(* IEC 61131-3 sources: daoli-st-library/DL_Process (part 7) *)

(* ---- FB_DL_SplicerAutoJoint.st ---- *)
//==============================================================================
// 功能块：FB_DL_SplicerAutoJoint ｜ 中文名称：自动接膜零停机顺控
// 所属子库：DL_Process ｜ 版本：v1.1.1 ｜ 兼容：CODESYS V3.5+ / TwinCAT 3 / 汇川 InoProShop
// 功能描述：卷材设备自动接膜（零停机换卷）顺控：旧卷余量预警 → 新卷预加速 → 速度同步
//           确认（容差 + 保持时长双条件）→ 裁切压合 → 尾料处理 → 回到监测相。
//           安全铁律：未同步绝不裁切——速度差超容差或保持时长不足时裁切一律挂起，宁可
//           等，不裁切（拉断料带的代价远高于停一拍）。余量按面积（卷径平方）比例折算，
//           按直径线性折算会把余量算大一倍以上（量纲教训：卷材体积随直径平方变化）。
//           本件只发预加速/裁切指令与状态，不驱动伺服、不控气阀（执行器归设备层）。
// 开源溯源 (Origin)：道莅 clean-room 防御性实现（原创，参考 公开工程惯例 分类与参数域）
// 单位表：卷径/芯径/满卷直径[mm] / 线速度[米每分] / 余量与预警门限[百分数] /
//         同步容差[百分数] / 时间窗[ms] / 扫描间隔[ms] / 接膜次数[次]
// 错误码表：16#0005_040A 信息级（余量预警触发，上升沿一次，不置 bError）/
//           16#0005_040B 信息级（同步窗未达，裁切挂起，不置 bError）/ 16#0005_0351
//           故障级（预加速超时中止且不裁切；兼「卷径组态非法（满卷直径 ≤ 芯径）」组态
//           分支，映射见本行反证句）/ 16#0005_0352 故障级（胶带未就绪或刀未归零，禁止
//           接膜，置 bError + 撤全部指令）/ 16#0005_0353 故障级（输入非有限，以及状态机
//           ELSE 非法状态兜底）。0351 共用反证句：组态非法、预加速超时与同步相超时
//           （v1.1.0 新增）在现有输出组合下不可观测出差异（均为 bError + bPreAccelCmd 撤
//           + bCutCmd 撤 + bSyncOk 撤 + bValid 撤），同步超时另由 bSyncTimeout 单拍事件可区分观测；
//           §4.17 亦明示组态分支映射入 0351，故共用不越段。0353 共用反证句：非有限
//           输入与非法状态在输出上同为全撤 + bError + eFault，不可观测出差异，故共用。
// 状态机：E_DL_SplicerState（eIdle=0 待机 / eMonitor=10 余量监测 / ePreAccel=20 新卷
//           预加速 / eSyncWait=30 同步确认 / eJointing=40 裁切压合 / eFault=99 故障兜底），
//           CASE 含 ELSE 兜底，ELSE 置 0353 且撤全部指令、许可撤。
// 边界行为：① 余量按面积比例 ((D^2 − core^2)/(full^2 − core^2)) x 100，D 低于芯径钳 0、
//           高于满卷钳 100；② fFullDiaMm <= fCoreDiaMm → 故障 0351 组态分支（分母为零
//           会产出伪余量，先判后算）；③ 预加速超 tPreAccelMax → 故障 0351 + 中止且绝不
//           裁切（停机保料优于拉断）；④ 同步未达（速度差 > 容差，或保持不足 tSyncHold）
//           → 裁切挂起 + 信息 040B（安全侧：宁可等，不裁切）；⑤ bTapeOk 或 bKnifeHome
//           为 FALSE → 禁止接膜 + 故障 0352；⑥ bStop → 中止并回 eIdle（同③不裁切）；
//           ⑦ 余量预警上升沿 → 信息 040A（用沿检测，防每拍刷屏）。
// 修订历史：v1.0.0 2026-11-17 首版（R25 派单 · §4.17）
//           v1.0.1 2026-11-17 终审补 eSyncWait 的「进相前置消失」第二退出条件（对外引脚契约零变更）：
//           bNewRollReady 撤销时退回 ePreAccel 相，由 tPreAccelMax 超时闸兜住，避免 bPreAccelCmd
//           长期拉住空卷（R98 家族）。两相 bCutCmd 均为 FALSE，「未同步绝不裁切」铁律不受影响。
//           v1.1.0 2026-11-17 R27 欠账收口（MINOR 升级，引脚契约只增不改、既有码位零变更）：
//           eSyncWait 相新增引脚 tSyncMax（同步等待超时，默认 T#5S）与自有计时器 fbTonSyncMax
//           （每周期无条件调用，仅 IN 条件化）；速度差持续超容差达 tSyncMax 即复用故障级 0351
//           （同段共用，反证句见错误码表 0351 行）并中止，bCutCmd 全程保持 FALSE；新增输出
//           bSyncTimeout（超时单拍事件，供审计计数）。
//           原挂账 R112 三要素收口：复现条件 = bNewRollReady 保持 TRUE 而速度差持续超容差（旧版将
//           无限期停在同步相）；禁用范围 = 无人值守连续线未配该超时者不得无人看管运行；修法取
//           ①新增 tSyncMax 引脚（默认 5 s 从紧口径）。
//           验收向量（VERSION 修订记录同步登记）：新卷就绪后速度差恒定 5%、容差 2% →
//           tSyncMax 之后置 0351、bSyncTimeout 单拍 TRUE、bCutCmd 全程 FALSE。
//           v1.1.1 2026-11-17 R27 终审修复（对外引脚与码位零变更）：fbTonSyncMax 的 IN 由
//           「eSyncWait AND NOT bSpeedWithin」改为「eSyncWait」按相驻留计时。原实现的看门狗
//           只在速度差超出容差时累积：速度差在容差边界抖动（模拟量噪声常态）时，同步超时
//           计时器与同步保持计时器交替复位，两者永不完成 → 相内无限滞留、段 8B 永不触发，
//           bPreAccelCmd 长期拉住空卷，恰是 v1.1.0 要收口的故障模式在抖动输入下的复现。
//           改为按相驻留计时后，相内总等待时长有上界，抖动亦能收口；正常同步（远早于
//           tSyncMax 完成）行为不变。验收向量：速度差在 2% 容差上下逐拍抖动 → tSyncMax 后 0351。
//==============================================================================
(*------------------------------------------------------------------------------
 * 枚举: E_DL_SplicerState（归属 DL_Process，与 FB_DL_SplicerAutoJoint 同文件）
 *----------------------------------------------------------------------------*)
TYPE E_DL_SplicerState :
(
    eIdle     := 0,   // 待机：指令全撤 / Idle, every command dropped
    eMonitor  := 10,  // 余量监测：算余量、报预警 / Monitoring the remaining roll
    ePreAccel := 20,  // 预加速：新卷升速，等就绪与同步 / Pre-accelerating the new roll
    eSyncWait := 30,  // 同步确认：速度差在容差内且保持达时 / Confirming the speed match
    eJointing := 40,  // 裁切压合：出裁切指令并在接膜窗内完成 / Cutting and joining
    eFault    := 99   // 故障兜底：超时/胶带刀具不就绪/非有限/非法状态 / Fault fallback
);
END_TYPE

(*==============================================================================
 * 功能块: FB_DL_SplicerAutoJoint
 * 调用约定: 每个扫描周期无条件调用一次；uDeltaTimeMs 必须注入真实任务间隔。
 *============================================================================*)
FUNCTION_BLOCK FB_DL_SplicerAutoJoint
VAR_INPUT
    fUnwindDiaMm    : LREAL;                       // 旧卷当前卷径 [mm] / Current unwinding roll diameter [mm]
    fCoreDiaMm      : LREAL;                       // 芯径 [mm]，须 > 0 / Core diameter [mm], must be > 0
    fFullDiaMm      : LREAL;                       // 满卷直径 [mm]，须 > 芯径 / Full roll diameter [mm], must exceed the core
    fWebSpeedMpm    : LREAL;                       // 旧卷线速度 [米每分] / Current web speed [m per min]
    fNewRollSpeedMpm : LREAL;                      // 新卷表面线速度 [米每分] / New roll surface speed [m per min]
    fRemainWarnPct  : LREAL := 15.0;               // 余量预警门限 [百分数] / Remaining-roll warning threshold [percent]
    fSyncTolPct     : LREAL := 2.0;                // 速度同步容差 [百分数] / Speed match tolerance [percent]
    tSyncHold       : TIME := T#500MS;             // 同步保持确认时长 [ms] / Speed match hold time [ms]
    tPreAccelMax    : TIME := T#20S;               // 预加速超时 [ms] / Pre-acceleration timeout [ms]
    tJointMax       : TIME := T#5S;                // 接膜（裁切压合）窗 [ms] / Joint window [ms]
    tSyncMax        : TIME := T#5S;                // 同步等待超时 [ms]，默认 5 s（eSyncWait 自有看门狗，小于 1 s 钳 1 s）/ Sync wait timeout [ms]
    bNewRollReady   : BOOL;                        // 新卷就绪（装卷到位、气路正常）/ New roll ready
    bKnifeHome      : BOOL;                        // 切刀在零位 / Knife at home position
    bTapeOk         : BOOL;                        // 胶带就绪 / Tape ready
    bStart          : BOOL;                        // 启动（取上升沿）/ Start, rising edge
    bStop           : BOOL;                        // 停止（中止并回待机，绝不裁切）/ Stop, aborts without cutting
    bReset          : BOOL;                        // 复位，上升沿回待机并清故障 / Reset, rising edge returns to idle
    uDeltaTimeMs    : UDINT;                       // 扫描间隔 [ms]，调用方注入，禁系统时间函数 / Scan interval [ms], caller-injected
END_VAR
VAR_OUTPUT
    bWarnLowRoll    : BOOL;                        // 余量预警（电平）/ Low-roll warning, level
    bPreAccelCmd    : BOOL;                        // 新卷预加速指令 / Pre-acceleration command
    bSyncOk         : BOOL;                        // 速度同步确认（容差 + 保持时长双条件）/ Speed match confirmed
    bSyncTimeout    : BOOL;                        // 同步超时事件（单拍脉冲，v1.1.0 新增）/ Sync-timeout event, single-scan pulse
    bCutCmd         : BOOL;                        // 裁切指令（未同步绝不为 TRUE）/ Cut command, never TRUE unless matched
    bJointDone      : BOOL;                        // 接膜完成（单拍脉冲）/ Joint completed, single-scan pulse
    fRemainPct      : LREAL;                       // 旧卷余量 [百分数]，按面积比例 / Remaining roll [percent], by area ratio
    uJointCount     : UDINT;                       // 接膜次数 [次]，饱和 / Joint count [pcs], saturating
    eErr            : UDINT;                       // 错误码，0 = 无错，码位 16#0005_040A 起信息级、16#0005_0351 起故障级（分带见错误码表） / Error code, 0 = no error, band info/fault per the code table
    bError          : BOOL;                        // 故障级标志，仅故障级错误置位 / Fault-class flag, set only on fault-level codes
    bValid          : BOOL;                        // 状态输出可用标志，失能/故障闸显式 FALSE / Status usable flag, explicit FALSE on disable/fault gates
    eState          : E_DL_SplicerState;           // 主状态机当前状态 / Current state of the main state machine
END_VAR
VAR
    fbReset         : R_TRIG;                      // 复位上升沿检测实例 / Reset rising edge detector
    fbStart         : R_TRIG;                      // 启动上升沿检测实例 / Start rising edge detector
    fbWarn          : R_TRIG;                      // 余量预警上升沿检测实例 / Low-roll warning rising edge detector
    fbTonPreAccel   : TON;                         // 预加速超时定时器实例 / Pre-acceleration timeout timer
    fbTonSyncHold   : TON;                         // 同步保持定时器实例 / Speed match hold timer
    fbTonJoint      : TON;                         // 接膜窗定时器实例 / Joint window timer
    fbTonSyncMax    : TON;                         // 同步相自有超时定时器实例（每周期无条件调用）/ Sync-phase watchdog timer instance
    tSyncMaxUse     : TIME;                        // 生效同步超时（下限钳 1 s 防误配置）/ Effective sync timeout, floored at 1 s
    fCoreSqMm2      : LREAL;                       // 芯径平方 [平方毫米] / Core diameter squared [mm2]
    fFullSqMm2      : LREAL;                       // 满卷直径平方 [平方毫米] / Full diameter squared [mm2]
    fDenomMm2       : LREAL;                       // 面积分母（满卷平方 − 芯径平方）[平方毫米] / Area denominator [mm2]
    fRemainNumMm2   : LREAL;                       // 面积分子（当前平方 − 芯径平方）[平方毫米] / Area numerator [mm2]
    fSpeedDiffPct   : LREAL;                       // 新旧卷速度差 [百分数] / Speed difference [percent]
    fTolEffPct      : LREAL;                       // 生效同步容差 [百分数] / Effective sync tolerance [percent]
    fWarnEffPct     : LREAL;                       // 生效预警门限 [百分数] / Effective warning threshold [percent]
    bNonFin         : BOOL;                        // 非有限判定中间标志 / Non-finite detection intermediate flag
    bSpeedWithin    : BOOL;                        // 速度差在容差内（瞬时）/ Speed difference within tolerance, instantaneous
    bJointOk        : BOOL;                        // 胶带与刀具均就绪 / Tape and knife both ready
    bFirstScan      : BOOL := TRUE;                // 上电首拍标志 / First-scan flag
END_VAR
VAR CONSTANT
    DL_SPJ_CODE_INFO_1 : UDINT := 16#0005_040A;    // 信息级槽 1（余量预警触发） / info slot 1
    DL_SPJ_CODE_INFO_2 : UDINT := 16#0005_040B;    // 信息级槽 2（同步窗未达，裁切挂起） / info slot 2
    DL_SPJ_CODE_FLT_1  : UDINT := 16#0005_0351;    // 故障级槽 1（预加速超时/卷径组态非法） / fault slot 1
    DL_SPJ_CODE_FLT_2  : UDINT := 16#0005_0352;    // 故障级槽 2（胶带未就绪/刀未归零） / fault slot 2
    DL_SPJ_CODE_FLT_3  : UDINT := 16#0005_0353;    // 故障级槽 3（非有限/非法状态兜底） / fault slot 3
    DL_SPJ_CNT_MAX     : UDINT := 16#FFFF_FFFE;    // 接膜计数饱和值 [次] / Joint counter saturation
    DL_SPJ_PCT         : LREAL := 100.0;           // 百分数系数 [百分数] / Percent factor
    DL_SPJ_ZERO        : LREAL := 0.0;             // 零值常量，避免裸字面量 [—] / Zero constant, avoids a bare literal
    DL_SPJ_TOL         : LREAL := 1.0E-6;          // 浮点比较容差 [—] / Float comparison tolerance
    DL_SPJ_INF         : LREAL := 1.7976931348623157E308; // LREAL 幅值上限，Inf 判据 / LREAL magnitude ceiling
END_VAR

(*------------------------------------------------------------------------------
 * 段 1｜无条件刷新区（红线 5）：三条沿检测与三个定时器在任意分支之外周期调用；
 *       定时器 IN 取上拍状态（单拍滞后对秒级时间窗无影响），计时链永不断流
 *----------------------------------------------------------------------------*)
bJointDone := FALSE;                               // 接膜完成为单拍脉冲，逐拍先清 / single-scan pulse cleared first
bSyncTimeout := FALSE;                             // 同步超时为单拍事件，逐拍先清 / sync-timeout event cleared first
tSyncMaxUse := tSyncMax;                           // 生效超时取引脚值 / effective timeout from the pin
IF tSyncMaxUse < T#1S THEN
    tSyncMaxUse := T#1S;                           // 超时下限钳 1 s（防 0 配置入相同拍误报）/ floored at 1 s
END_IF
fbReset(CLK := bReset);                            // 复位沿检测无条件刷新 / reset edge refreshed unconditionally
fbStart(CLK := bStart);                            // 启动沿检测无条件刷新 / start edge refreshed unconditionally
fbTonPreAccel(IN := (eState = E_DL_SplicerState.ePreAccel), PT := tPreAccelMax);   // 预加速超时计时 / pre-acceleration timeout
fbTonSyncHold(IN := (eState = E_DL_SplicerState.eSyncWait) AND bSpeedWithin, PT := tSyncHold);   // 同步保持计时 / speed match hold
fbTonJoint(IN := (eState = E_DL_SplicerState.eJointing), PT := tJointMax);         // 接膜窗计时 / joint window
fbTonSyncMax(IN := (eState = E_DL_SplicerState.eSyncWait), PT := tSyncMaxUse);   // v1.1.1 改为按相驻留计时（见修订史 R27-3）/ sync watchdog on phase residency
fbWarn(CLK := bWarnLowRoll);                       // 预警上升沿检测无条件刷新 / warning edge refreshed unconditionally

(*------------------------------------------------------------------------------
 * 段 2｜复位沿处理（改写置于沿后，防吞沿 R39）
 *----------------------------------------------------------------------------*)
IF fbReset.Q THEN
    eState := E_DL_SplicerState.eIdle;
    eErr   := 0;                        // 复位清码 / reset clears the code
    bError := FALSE;                               // 复位清故障 / reset clears the fault
    bPreAccelCmd := FALSE;                         // 预加速指令撤 / pre-acceleration dropped
    bCutCmd := FALSE;                              // 裁切指令撤 / cut command dropped
    bSyncOk := FALSE;                              // 同步确认撤 / sync confirmation dropped
    bFirstScan := TRUE;                            // 重新首拍化 / re-initialize first scan
END_IF

(*------------------------------------------------------------------------------
 * 段 3｜非有限输入闸：映射入 0353（与非法状态共用，反证句见错误码表）
 *       安全侧：撤全部指令，绝不裁切
 *----------------------------------------------------------------------------*)
bNonFin := (fUnwindDiaMm <> fUnwindDiaMm) OR (ABS(fUnwindDiaMm) >= DL_SPJ_INF)
        OR (fCoreDiaMm <> fCoreDiaMm) OR (ABS(fCoreDiaMm) >= DL_SPJ_INF)
        OR (fFullDiaMm <> fFullDiaMm) OR (ABS(fFullDiaMm) >= DL_SPJ_INF)
        OR (fWebSpeedMpm <> fWebSpeedMpm) OR (ABS(fWebSpeedMpm) >= DL_SPJ_INF)
        OR (fNewRollSpeedMpm <> fNewRollSpeedMpm) OR (ABS(fNewRollSpeedMpm) >= DL_SPJ_INF)
        OR (fRemainWarnPct <> fRemainWarnPct) OR (ABS(fRemainWarnPct) >= DL_SPJ_INF)
        OR (fSyncTolPct <> fSyncTolPct) OR (ABS(fSyncTolPct) >= DL_SPJ_INF);   // 引脚非有限汇总 / pins non-finite
IF bNonFin THEN
    eState := E_DL_SplicerState.eFault;            // 进故障相 / enter fault state
    eErr   := DL_SPJ_CODE_FLT_3;                   // 故障级：输入非有限 / fault: non-finite input
    bError := TRUE;                                // 故障级必置 bError（R45 配对）/ fault-class pairs with bError
    bValid := FALSE;                               // 状态不可用 / status unusable
    bPreAccelCmd := FALSE;                         // 预加速指令撤 / pre-acceleration dropped
    bCutCmd := FALSE;                              // 裁切指令撤（安全侧：绝不裁切）/ cut dropped, never cut
    bSyncOk := FALSE;                              // 同步确认撤 / sync confirmation dropped
    RETURN;
END_IF

(*------------------------------------------------------------------------------
 * 段 4｜卷径组态闸：满卷直径必须严格大于芯径（否则面积分母为零，余量必假）
 *       §4.17 明示本组态分支映射入 0351
 *----------------------------------------------------------------------------*)
IF (fCoreDiaMm <= DL_SPJ_TOL) OR (fFullDiaMm <= fCoreDiaMm + DL_SPJ_TOL) THEN
    eState := E_DL_SplicerState.eFault;            // 进故障相 / enter fault state
    eErr   := DL_SPJ_CODE_FLT_1;                   // 故障级：卷径组态非法（映射入 0351）/ fault: roll diameter configuration invalid
    bError := TRUE;                                // 故障级必置 bError（R45 配对）/ fault-class pairs with bError
    bValid := FALSE;                               // 状态不可用 / status unusable
    bPreAccelCmd := FALSE;                         // 预加速指令撤 / pre-acceleration dropped
    bCutCmd := FALSE;                              // 裁切指令撤安全侧 / cut dropped, safe side
    bSyncOk := FALSE;                              // 同步确认撤 / sync confirmation dropped
    fRemainPct := DL_SPJ_ZERO;                     // 余量不可算，输出 0 而不是伪值 / remaining reported as 0, not a fake value
    RETURN;
END_IF

(*------------------------------------------------------------------------------
 * 段 5｜余量面积比例折算：((D^2 − core^2) / (full^2 − core^2)) x 100
 *       按直径线性折算会把余量算大一倍以上（面积随直径平方变化，R12 同族量纲教训）
 *----------------------------------------------------------------------------*)
fCoreSqMm2 := fCoreDiaMm * fCoreDiaMm;             // 芯径平方 [平方毫米] / core squared [mm2]
fFullSqMm2 := fFullDiaMm * fFullDiaMm;             // 满卷直径平方 [平方毫米] / full squared [mm2]
fDenomMm2 := fFullSqMm2 - fCoreSqMm2;              // 面积分母（段 4 已保证为正）[平方毫米] / area denominator, proven positive
fRemainNumMm2 := (fUnwindDiaMm * fUnwindDiaMm) - fCoreSqMm2;   // 面积分子 [平方毫米] / area numerator [mm2]
IF fRemainNumMm2 < DL_SPJ_ZERO THEN
    fRemainNumMm2 := DL_SPJ_ZERO;                  // 卷径低于芯径：分子钳零（欠卷异常不产出负余量）/ numerator floored at zero
END_IF
fRemainPct := fRemainNumMm2 / fDenomMm2 * DL_SPJ_PCT;   // 余量 [百分数] / remaining [percent]
IF fRemainPct > DL_SPJ_PCT THEN
    fRemainPct := DL_SPJ_PCT;                      // 卷径超满卷：钳 100 / clamped to 100
END_IF
IF fRemainPct < DL_SPJ_ZERO THEN
    fRemainPct := DL_SPJ_ZERO;                     // 下限防护 / floor guard
END_IF
fWarnEffPct := fRemainWarnPct;                     // 预警门限工作副本 [百分数] / warning threshold working copy
IF fWarnEffPct < DL_SPJ_ZERO THEN
    fWarnEffPct := DL_SPJ_ZERO;                    // 门限下限钳位 / threshold floored
END_IF
IF fWarnEffPct > DL_SPJ_PCT THEN
    fWarnEffPct := DL_SPJ_PCT;                     // 门限上限钳位 / threshold clamped to 100
END_IF
bWarnLowRoll := (fRemainPct <= fWarnEffPct);       // 余量预警（电平）/ low-roll warning, level

(*------------------------------------------------------------------------------
 * 段 6｜速度同步判据：|旧卷 − 新卷| / 旧卷 x 100 <= 容差（除子先判零，低速记不同步）
 *----------------------------------------------------------------------------*)
fTolEffPct := fSyncTolPct;                         // 容差工作副本 [百分数] / tolerance working copy
IF fTolEffPct < DL_SPJ_ZERO THEN
    fTolEffPct := DL_SPJ_ZERO;                     // 负容差钳零（等价于要求完全相等）/ negative tolerance floored
END_IF
IF fWebSpeedMpm > DL_SPJ_TOL THEN
    fSpeedDiffPct := ABS(fWebSpeedMpm - fNewRollSpeedMpm) / fWebSpeedMpm * DL_SPJ_PCT;   // 速度差 [百分数] / speed difference [percent]
    bSpeedWithin := (fSpeedDiffPct <= fTolEffPct); // 容差内判据 / within-tolerance predicate
ELSE
    fSpeedDiffPct := DL_SPJ_PCT;                   // 旧卷静止：速度差按满刻度记（不可判即不同步）/ web at standstill, treated as not matched
    bSpeedWithin := FALSE;                         // 静止时不允许裁切 / no cut while the web stands still
END_IF
bJointOk := bTapeOk AND bKnifeHome;                // 胶带与刀具就绪判据 / tape and knife ready predicate
bSyncOk := bSpeedWithin AND fbTonSyncHold.Q AND (eState = E_DL_SplicerState.eSyncWait);   // 同步确认＝容差内且保持达时 / match confirmed

(*------------------------------------------------------------------------------
 * 段 7｜禁止接膜闸：胶带未就绪或刀未归零 → 0352 + 撤指令（不裁切）
 *----------------------------------------------------------------------------*)
IF (NOT bJointOk) AND ((eState = E_DL_SplicerState.ePreAccel) OR (eState = E_DL_SplicerState.eSyncWait)
                       OR (eState = E_DL_SplicerState.eJointing)) THEN
    eState := E_DL_SplicerState.eFault;            // 进故障相 / enter fault state
    eErr   := DL_SPJ_CODE_FLT_2;                   // 故障级：胶带未就绪/刀未归零，禁止接膜 / fault: tape or knife not ready
    bError := TRUE;                                // 故障级必置 bError（R45 配对）/ fault-class pairs with bError
    bValid := FALSE;                               // 状态不可用 / status unusable
    bPreAccelCmd := FALSE;                         // 预加速指令撤 / pre-acceleration dropped
    bCutCmd := FALSE;                              // 裁切指令撤（禁止接膜）/ cut dropped, joining forbidden
    bSyncOk := FALSE;                              // 同步确认撤 / sync confirmation dropped
    RETURN;
END_IF

(*------------------------------------------------------------------------------
 * 段 8｜预加速超时闸：0351 + 中止且绝不裁切（停机保料优于拉断）
 *----------------------------------------------------------------------------*)
IF (eState = E_DL_SplicerState.ePreAccel) AND fbTonPreAccel.Q THEN
    eState := E_DL_SplicerState.eFault;            // 进故障相 / enter fault state
    eErr   := DL_SPJ_CODE_FLT_1;                   // 故障级：预加速超时，中止且不裁切 / fault: pre-acceleration timeout, abort without cutting
    bError := TRUE;                                // 故障级必置 bError（R45 配对）/ fault-class pairs with bError
    bValid := FALSE;                               // 状态不可用 / status unusable
    bPreAccelCmd := FALSE;                         // 预加速指令撤 / pre-acceleration dropped
    bCutCmd := FALSE;                              // 裁切指令撤（绝不裁切）/ cut dropped, never cut
    bSyncOk := FALSE;                              // 同步确认撤 / sync confirmation dropped
    RETURN;
END_IF

(*------------------------------------------------------------------------------
 * 段 8B｜同步相超时闸（v1.1.0 欠账收口，R112 家族）：速度差持续超容差达 tSyncMax
 *       → 复用故障级 0351 并中止，bCutCmd 全程 FALSE（安全铁律：未同步绝不裁切）
 *----------------------------------------------------------------------------*)
IF (eState = E_DL_SplicerState.eSyncWait) AND fbTonSyncMax.Q THEN
    eState := E_DL_SplicerState.eFault;            // 进故障相 / enter fault state
    eErr   := DL_SPJ_CODE_FLT_1;                   // 故障级：同步超时（与预加速超时同段共用，反证句见头注）/ fault: sync timeout
    bError := TRUE;                                // 故障级必置 bError（R45 配对）/ fault-class pairs with bError
    bValid := FALSE;                               // 状态不可用 / status unusable
    bPreAccelCmd := FALSE;                         // 预加速指令撤 / pre-acceleration dropped
    bCutCmd := FALSE;                              // 裁切指令撤（绝不裁切）/ cut dropped, never cut
    bSyncOk := FALSE;                              // 同步确认撤 / sync confirmation dropped
    bSyncTimeout := TRUE;                          // 同步超时单拍事件 / single-scan sync-timeout event
    RETURN;
END_IF

(*------------------------------------------------------------------------------
 * 段 9｜状态机：CASE 含 ELSE 兜底（非法状态 → 0353 + 撤全部指令 + 许可撤）
 *----------------------------------------------------------------------------*)
CASE eState OF

    E_DL_SplicerState.eIdle:
        bPreAccelCmd := FALSE;                     // 待机预加速撤 / pre-acceleration dropped in idle
        bCutCmd := FALSE;                          // 待机裁切撤 / cut dropped in idle
        bSyncOk := FALSE;                          // 待机同步确认撤 / sync confirmation dropped in idle
        bValid := FALSE;                           // 失能闸显式不可用（R72）/ explicit FALSE on the disable gate
        eErr := 0;                      // 待机无错 / no error in idle
        bError := FALSE;                           // 待机无故障 / no fault in idle
        IF fbStart.Q THEN
            IF bJointOk THEN
                eState := E_DL_SplicerState.ePreAccel;   // 就绪才允许预加速 / pre-acceleration only when ready
                bFirstScan := FALSE;               // 首拍标志清除 / first-scan flag cleared
            ELSE
                eState := E_DL_SplicerState.eFault;      // 不就绪直接进故障相（0352）/ not ready enters the fault state
                eErr := DL_SPJ_CODE_FLT_2;         // 故障级：胶带未就绪/刀未归零 / fault: tape or knife not ready
                bError := TRUE;                    // 故障级必置 bError（R45 配对）/ fault-class pairs with bError
            END_IF
        ELSE
            eState := E_DL_SplicerState.eMonitor;  // 无启动沿：进常驻余量监测相（监测是被动功能，无需启动）/ passive monitoring needs no start
        END_IF

    E_DL_SplicerState.eMonitor:
        bPreAccelCmd := FALSE;                     // 监测相不预加速 / no pre-acceleration while monitoring
        bCutCmd := FALSE;                          // 监测相不裁切 / no cut while monitoring
        bSyncOk := FALSE;                          // 监测相无同步确认 / no sync confirmation while monitoring
        bValid := TRUE;                            // 余量与预警可用 / remaining and warning usable
        bError := FALSE;                           // 监测相无故障 / no fault while monitoring
        IF fbWarn.Q THEN
            eErr := DL_SPJ_CODE_INFO_1;            // 信息级：余量预警触发（上升沿一次）/ info: low-roll warning, once per rising edge
        ELSE
            eErr := 0;                  // 非预警沿不占码位 / no code without a warning edge
        END_IF
        IF fbStart.Q AND bJointOk THEN
            eState := E_DL_SplicerState.ePreAccel; // 启动且就绪进预加速 / start with readiness enters pre-acceleration
        ELSIF fbStart.Q AND (NOT bJointOk) THEN
            eState := E_DL_SplicerState.eFault;    // 启动但不就绪：禁止接膜 / start without readiness forbids joining
            eErr := DL_SPJ_CODE_FLT_2;             // 故障级：胶带未就绪/刀未归零 / fault: tape or knife not ready
            bError := TRUE;                        // 故障级必置 bError（R45 配对）/ fault-class pairs with bError
            bValid := FALSE;                       // 状态不可用 / status unusable
        END_IF

    E_DL_SplicerState.ePreAccel:
        bPreAccelCmd := TRUE;                      // 新卷预加速指令 / pre-acceleration command
        bCutCmd := FALSE;                          // 预加速相绝不裁切 / never cut while pre-accelerating
        bSyncOk := FALSE;                          // 预加速相尚无同步确认 / not yet confirmed
        bValid := TRUE;                            // 状态可用 / status usable
        bError := FALSE;                           // 本相无故障（超时已由段 8 处置）/ no fault here, timeout handled earlier
        eErr := 0;                      // 预加速相先清码 / clear the code first
        IF bNewRollReady THEN
            eState := E_DL_SplicerState.eSyncWait; // 新卷就绪进同步确认 / new roll ready enters the sync wait
        END_IF

    E_DL_SplicerState.eSyncWait:
        bPreAccelCmd := TRUE;                      // 预加速保持（同步需要维持速度）/ pre-acceleration held to keep the speed
        bCutCmd := FALSE;                          // 未确认绝不出裁切 / no cut before confirmation
        bValid := TRUE;                            // 状态可用 / status usable
        bError := FALSE;                           // 本相无故障 / no fault here
        IF bSyncOk THEN
            eErr := 0;                  // 已同步：无提示 / matched, no hint
            bCutCmd := TRUE;                       // 同步确认后才出裁切指令 / cut only after the match is confirmed
            eState := E_DL_SplicerState.eJointing; // 进裁切压合相 / enter cutting and joining
        ELSIF NOT bNewRollReady THEN
            // v1.0.1 补「进相前置消失」退出条件（R98 家族第二出口）：新卷预加速/就绪条件撤销时，
            // 本相已失去同步对象，继续滞留只会让 bPreAccelCmd 长期拉住空卷。退回 ePreAccel 相，
            // 由该相的 tPreAccelMax 超时闸兜住（仍保持「绝不裁切」——两相 bCutCmd 均为 FALSE）。
            eErr := DL_SPJ_CODE_INFO_2;            // 信息级：仍报同步未达 / info: still not matched
            eState := E_DL_SplicerState.ePreAccel; // 退回预加速相（前置消失退出条件）/ back to pre-acceleration, precondition gone
        ELSE
            eErr := DL_SPJ_CODE_INFO_2;            // 信息级：同步窗未达，裁切挂起（宁可等，不裁切）/ info: cut suspended
        END_IF

    E_DL_SplicerState.eJointing:
        bCutCmd := TRUE;                           // 裁切指令保持（接膜窗内）/ cut command held inside the joint window
        bPreAccelCmd := TRUE;                      // 预加速保持到接膜完成 / pre-acceleration held until the joint completes
        bValid := TRUE;                            // 状态可用 / status usable
        bError := FALSE;                           // 本相无故障 / no fault here
        eErr := 0;                      // 接膜相无错 / no error while joining
        IF fbTonJoint.Q THEN
            bCutCmd := FALSE;                      // 接膜窗到点撤裁切 / cut dropped when the window elapses
            bPreAccelCmd := FALSE;                 // 预加速撤 / pre-acceleration dropped
            bJointDone := TRUE;                    // 接膜完成单拍脉冲 / single-scan joint-done pulse
            IF uJointCount < DL_SPJ_CNT_MAX THEN
                uJointCount := uJointCount + 1;    // 接膜次数饱和自增 [次] / saturating joint increment
            END_IF
            eState := E_DL_SplicerState.eMonitor;  // 回监测相监测新卷余量 / back to monitoring the new roll
        END_IF

    E_DL_SplicerState.eFault:
        bPreAccelCmd := FALSE;                     // 故障闸撤预加速（R72）/ pre-acceleration dropped on the fault gate
        bCutCmd := FALSE;                          // 故障闸撤裁切（绝不裁切）/ cut dropped, never cut
        bSyncOk := FALSE;                          // 同步确认撤 / sync confirmation dropped
        bValid := FALSE;                           // 故障闸显式不可用 / explicit FALSE on the fault gate
        bError := TRUE;                            // 故障级必置 bError（R45 配对）/ fault-class pairs with bError
        IF eErr = 0 THEN
            eErr := DL_SPJ_CODE_FLT_3;             // 入口无码时按非法状态兜底（R45：bError 必须有对应码）/ illegal-state fallback
        END_IF
        IF fbReset.Q THEN
            eState := E_DL_SplicerState.eIdle;     // 仅复位可退出故障相 / only reset leaves the fault state
        END_IF

    ELSE
        eState := E_DL_SplicerState.eFault;        // 非法状态兜底 / illegal-state fallback
        eErr := DL_SPJ_CODE_FLT_3;                 // 故障级兜底：非法状态 / fault fallback: illegal state
        bError := TRUE;                            // 故障级必置 bError（R45 配对）/ fault-class pairs with bError
        bValid := FALSE;                           // 状态不可用 / status unusable
        bPreAccelCmd := FALSE;                     // 预加速指令撤 / pre-acceleration dropped
        bCutCmd := FALSE;                          // 裁切指令撤安全侧（绝不裁切）/ cut dropped, never cut
        bSyncOk := FALSE;                          // 同步确认撤 / sync confirmation dropped

END_CASE

(*------------------------------------------------------------------------------
 * 段 10｜停止闸（电平，最后判，覆盖各相输出）：中止并回待机，绝不裁切。
 *       放在 CASE 之后是为了让「停止」压过任何相内指令（安全侧优先级最高）
 *----------------------------------------------------------------------------*)
IF bStop THEN
    eState := E_DL_SplicerState.eIdle;             // 回待机 / back to idle
    bPreAccelCmd := FALSE;                         // 预加速撤 / pre-acceleration dropped
    bCutCmd := FALSE;                              // 裁切撤（中止不裁切）/ cut dropped, abort without cutting
    bSyncOk := FALSE;                              // 同步确认撤 / sync confirmation dropped
    bValid := FALSE;                               // 停止闸显式不可用（R72）/ explicit FALSE on the stop gate
    bJointDone := FALSE;                           // 停止不产生完成脉冲 / no done pulse on a stop
END_IF
END_FUNCTION_BLOCK

(* ---- FB_DL_StretchWrapSeq.st ---- *)
(*==============================================================================
 * 组件名称 (Component)  : FB_DL_StretchWrapSeq
 * 所属子库 (Sublibrary) : DL_Process
 * 当前版本 (Version)    : 1.0.2
 * 兼容性   (Platform)   : CODESYS 3.5 / TwinCAT 3 / 汇川 InoProShop / Machine Expert
 *                         仅依赖 Standard.library（TON / R_TRIG），零厂商方言
 * 来源标签 (Source)     : t2-7-packml（工站最小子集范式，clean-room 编写）
 * 功能描述 (Function)   : 缠绕膜包装机七态最小顺控：预压 -> 底圈 -> 顶圈（圈数
 *                         配方：底 / 顶 / 总圈数三项）-> 切膜 -> 保持 -> 完成。
 *                         转盘旋转反馈经 R_TRIG 沿计数（计数饱和 255）；膜断检测
 *                         联锁暂停——暂停在圈数边界生效（当前圈转完即停），恢复
 *                         后从当前圈数继续（不重头，ISA-88 相语义次源）。
 * 范式互引 (Paradigm)   : 工站顺控范式参照 FB_DL_PickAndPlaceStation；PackML 17 态
 *                         全集属主为 FB_DL_PackMlStateMachine——本件刻意做七态
 *                         最小子集，全集语义（阻塞 / 中止 / 清空）归全集属主。
 * 边界与语义披露 (Boundary disclosure) :
 *   1) 圈数配方域 1..255：越界组态级故障拒绝启动（锁存至复位沿 + 配方改对）；
 *      总圈数与底 / 顶之和不一致为信息级（以底 + 顶之和为准执行）。
 *   2) 转盘反馈丢失超时锁存（故障级）：判据 = 驱动输出有效 AND 本拍无旋转沿，
 *      TON 逐段断输入（R40 家族口径）；解除 = 复位沿 AND 反馈恢复。
 *   3) 暂停双源（膜断检测 / 操作暂停请求）合并为同一暂停挂起位，在圈数边界
 *      生效：暂停挂起期间当前圈转完即停，驱动输出切断，圈数保持。
 *   4) 切膜失败出口（产品裁定，v1.0.2 点修②）：切膜重试计数饱和（nCutRetryMax 封顶
 *      不回绕）后**不再自动重切**——单次窗再次超时即判定切膜失败：置故障级码 +
 *      bCutFail 锁存 + 迁 eFault，切断 bCutOut 与转盘驱动，停机待人工处理；
 *      解除唯一路径为人工复位（bReset 上升沿 AND 配方合法），复位后回 eIdle 从头
 *      开始（重试计数在 eIdle 受理时清零，不延续失败票的计数）。
 *   5) 压膜释放口径（产品裁定，v1.0.2 点修⑦）：bPreClampOut 仅表达「预压建压」
 *      一个动作，只在 ePreClamp 相有效；一进入底圈段即释放，并在底 / 顶圈段
 *      **全程保持释放**（膜被转盘牵引缠绕，压膜件继续压住会压出膜皱 / 拉断），
 *      切膜 / 保持 / 空闲 / 故障相同样释放。释放由状态派生式结构性保证，
 *      不挂单拍标志、不由暂停位改写（暂停只在圈边界截停驱动，不改压膜）。
 *   6) eIdle 相执行输出清零（R57 LWF 家族扫描范式前置合规）。
 * 配比约束 (R100)       : tTurnLoss 须大于转盘单圈周期的 1.5 倍（防正常圈间隔误判）；
 *                         tCutTimeout > tCutDwell（切膜窗必须宽于重试间隔窗）。
 * 故障码表 (Error codes) :
 *   16#0005_03A9 [故障级] 圈数配方组态非法（<1 或 >255），拒绝启动
 *                 反证：拒绝启动与「未按启动」输出组合相同，码位唯一可见。
 *   16#0005_03AA [故障级] 转盘反馈丢失超时，锁存至复位沿 + 反馈恢复
 *                 反证：顺控停摆与暂停态输出组合相似但成因完全不同（机械 vs 操作），必须独立码位。
 *   16#0005_04D1 [信息级] 膜断检测触发，暂停挂起（事件流水归档）
 *                 反证：bPauseHold 已表达暂停态，但暂停双源（膜断 / 人工）不可区分。
 *   16#0005_04D2 [信息级] 总圈数与底 / 顶之和不一致，按底 + 顶之和执行
 *                 反证：不一致时执行结果与显式填一致值相同，无码不可区分。
 *   16#0005_04D3 [信息级] 切膜重试计数已饱和（封顶不回绕）
 *                 反证：饱和计数与恰好达上限计数输出相同，无码不可区分。
 *   16#0005_03B3 [故障级] 切膜失败（重试饱和后单次窗再次超时），停机待人工
 *                 反证：失败停机与「反馈丢失」同为 eFault + bError，但成因与处置
 *                 完全不同（反馈丢失复位后可从现场恢复；切膜失败必须人工拆膜）；
 *                 且原实现无出口时 eCut 永驻、bCutOut 常励磁，故障态与「切膜中」
 *                 输出组合无法区分（R190 归因唯一，R69 点修②）。
 * 码位总账 (Code ledger) : 16#0005_03A9 / 03AA / 03B3 用 ｜ 16#0005_04D1 / 04D2 / 04D3 用
 * 依赖     (Depends)    : 无 DL_ 内部依赖；Standard.library: TON / R_TRIG
 * 红线自检 (Redline)    : R1 ✓ 零全局变量与 VAR_EXTERNAL ｜ R2 ✓ 零 %I/%Q 物理地址
 *                         R3 ✓ 纯 IEC 61131-3 ｜ R4 ✓ 配方域闸 / 计数饱和 / 域闸全枚举
 *                         R5 ✓ 全变量中英双语同行注释 ｜ R6 ✓ 七态 ENUM + CASE + ELSE 兜底
 *                         R7 ✓ 四沿四计时主体最前部无条件刷新
 * 修订历史 (Revision)   :
 *   2026-11-22  v1.0.0  首版入库（R68 构建轮 · 批 3 · 目标 12）
 *   2026-11-22  v1.0.1  终审就地修④：总圈计数上限改用 510（原以单段上界 255 作总数闸，合法配方 >255 圈即死锁）
 *   2026-11-22  v1.0.2  R69 点修②：eCut 相补切膜失败出口（重试饱和后单次窗再超时 -> 03B3 +
 *                       bCutFail 锁存 + 迁 eFault 停机待人工，不自动重切，人工复位解除）；
 *                       点修⑦：bPreClampOut 语义固化（仅预压相有效，圈段全程释放防膜皱）
 *============================================================================*)

(*-----------------------------------------------------------------------------
 * 枚举: E_DL_WrapSeqState（归属 DL_Process，与 FB_DL_StretchWrapSeq 同文件）
 *----------------------------------------------------------------------------*)
TYPE E_DL_WrapSeqState :
(
    eIdle     := 0,    // 空闲：输出全清（R57 前置合规）/ Idle, all outputs cleared
    ePreClamp := 10,   // 预压：压膜建立 / Pre-clamp, film pressed
    eBottom   := 20,   // 底圈段：转盘计数 / Bottom turns, counting
    eTop      := 30,   // 顶圈段：转盘计数 / Top turns, counting
    eCut      := 40,   // 切膜：重试节流 / Film cut with retry throttle
    eDwell    := 50,   // 保持：保持窗计时 / Dwell window timing
    eFault    := 99    // 配方 / 反馈丢失 / 切膜失败 锁存 / Recipe, loss or cut failure latched
);
END_TYPE

(*==============================================================================
 * 功能块: FB_DL_StretchWrapSeq
 * 调用约定: 每个扫描周期无条件调用一次。
 *============================================================================*)
FUNCTION_BLOCK FB_DL_StretchWrapSeq
VAR_INPUT
    bStartCmd    : BOOL;                 // 启动命令（上升沿受理）/ Start command, rising edge accepted
    bStopCmd     : BOOL;                 // 停止命令（电平，任意相退出）/ Stop command, level, exits any phase
    bPauseReq    : BOOL;                 // 操作暂停请求（电平）/ Operator pause request, level
    bFilmBreak   : BOOL;                 // 膜断检测（电平，联锁暂停源）/ Film break detection, interlock pause source
    bTurnFb      : BOOL;                 // 转盘旋转反馈（每圈一脉冲）/ Turntable feedback, one pulse per revolution
    bPreClampFb  : BOOL;                 // 预压到位反馈 / Pre-clamp in-position feedback
    bCutDone     : BOOL;                 // 切膜完成反馈 / Film cut done feedback
    nBottomTurns : INT := 2;             // 底圈数配方 [圈]，域 1..255 / Bottom turns recipe
    nTopTurns    : INT := 3;             // 顶圈数配方 [圈]，域 1..255 / Top turns recipe
    nTotalTurns  : INT := 5;             // 总圈数配方 [圈]，仅一致性核对 / Total turns recipe, consistency only
    nCutRetryMax : INT := 3;             // 切膜重试上限 [次] / Film cut retry ceiling
    tPreClamp    : TIME := T#2S;         // 预压建压窗 [s] / Pre-clamp build-up window [s]
    tTurnLoss    : TIME := T#10S;        // 转盘反馈丢失超时 [s] / Turntable feedback loss timeout [s]
    tCutTimeout  : TIME := T#5S;         // 切膜单次窗 [s] / Film cut single window [s]
    tCutDwell    : TIME := T#1S;         // 切膜重试间隔窗 [s] / Film cut retry interval [s]
    tDwellHold   : TIME := T#3S;         // 保持窗时长 [s] / Dwell hold duration [s]
    bEnable      : BOOL := TRUE;         // 使能 / Enable
    bReset       : BOOL;                 // 上升沿：清配方 / 反馈丢失锁存 / Rising edge: clear latches
END_VAR
VAR_OUTPUT
    bTurnDrive  : BOOL;                  // 转盘驱动输出 / Turntable drive output
    bPreClampOut: BOOL;                  // 预压输出 / Pre-clamp output
    bCutOut     : BOOL;                  // 切膜输出 / Film cut output
    bPauseHold  : BOOL;                  // 暂停挂起（圈边界生效）/ Pause hold, effective at turn boundary
    bSeqActive  : BOOL;                  // 顺控进行中 / Sequence active
    bSeqDone    : BOOL;                  // 顺控完成脉冲（单拍）/ Sequence done pulse, single scan
    nTurnsDone  : INT;                   // 已完成总圈数 [圈] / Total turns completed
    nCutRetries : INT;                   // 切膜重试计数 [次]，饱和 / Film cut retries, saturating
    bCutFail    : BOOL;                  // 切膜失败锁存（停机待人工，人工复位解除）/ Cut failure latch, cleared by manual reset
    bError      : BOOL;                  // 故障标志（配方 / 反馈丢失）/ Fault flag
    uErrorId    : UDINT;                 // 故障码，0 = 无故障 / Error code, 0 = none
    eState      : E_DL_WrapSeqState;     // 当前状态（供 HMI 诊断）/ Current state
END_VAR
VAR
    fbTrigStart  : R_TRIG;               // 启动沿检测实例 / Start edge detector
    fbTrigReset  : R_TRIG;               // 复位沿检测实例 / Reset edge detector
    fbTrigFilm   : R_TRIG;               // 膜断沿检测实例（事件码用）/ Film break edge detector
    rTrigTurn    : R_TRIG;               // 转盘圈脉冲沿计数实例 / Turn pulse counting edge
    tonPre       : TON;                  // 预压建压计时实例 / Pre-clamp timer
    tonTurnLoss  : TON;                  // 转盘反馈丢失计时实例 / Turntable loss timer
    tonCutTo     : TON;                  // 切膜单次窗计时实例 / Film cut window timer
    tonCutDwell  : TON;                  // 切膜重试间隔窗（自复位）实例 / Retry interval timer, self resetting
    tonDwellHold : TON;                  // 保持窗计时实例 / Dwell hold timer
    eStateInt    : E_DL_WrapSeqState;    // 主状态机内部当前态 / Internal state machine state
    nBottomDone  : INT;                  // 底圈已完成圈数 [圈] / Bottom turns completed
    nTopDone     : INT;                  // 顶圈已完成圈数 [圈] / Top turns completed
    nRetryInt    : INT;                  // 切膜重试计数内部副本 / Internal retry count
    bPausePend   : BOOL;                 // 暂停挂起请求（双源合并）/ Pause pending, dual source merged
    bPauseHoldInt: BOOL;                 // 暂停边界生效保持位 / Pause hold latched at boundary
    bRecipeBad   : BOOL;                 // 本拍配方组态非法 / Recipe illegal this scan
    bRecipeLatch : BOOL;                 // 配方故障锁存（复位沿清除）/ Recipe fault latch
    bTotalDiff   : BOOL;                 // 总圈数与底 / 顶之和不一致 / Total mismatch with the sum
    bTurnLossInt : BOOL;                 // 反馈丢失锁存内部副本 / Internal feedback loss latch
    bCutFailInt  : BOOL;                 // 切膜失败锁存内部副本（人工复位解除）/ Internal cut failure latch
    bDoneT       : BOOL;                 // 完成脉冲内部副本（单拍）/ Internal done pulse copy
    bTurnDriveInt: BOOL;                 // 驱动输出内部派生 / Internal drive output derivation
    bErrorInt    : BOOL;                 // 本拍故障置位累加（出口归并）/ Fault set accumulator
    bFirstScan   : BOOL := TRUE;         // 上电首扫标志 / First-scan flag
END_VAR
VAR CONSTANT
    DL_WR_TURNS_MAX : INT := 255;    // 单段圈数上限 [圈]（配方域上界）/ Turns ceiling per recipe
    DL_WR_TOTAL_MAX : INT := 510;    // 总圈数上限 [圈]（= 2 x 单段上界，终审就地修 v1.0.1）/ Total turns ceiling
    DL_WR_RETRY_MAX : INT := 8;      // 重试计数硬饱和 [次]（防 INT 溢出兜底）/ Retry hard saturation
END_VAR

(*------------------------------------------------------------------------------
 * 段 1｜无条件刷新区（红线 R7）：四沿五计时全部位于主体最前部
 *      Unconditional refresh: four edges and five timers at the very top
 *      计时器 IN 全部为内部派生量（R40 断输入口径）
 *-----------------------------------------------------------------------------*)
fbTrigStart(CLK := bStartCmd);
fbTrigReset(CLK := bReset);
fbTrigFilm(CLK := bFilmBreak);
rTrigTurn(CLK := bTurnFb);

tonPre(IN := (eStateInt = E_DL_WrapSeqState.ePreClamp) AND (NOT bPreClampFb), PT := tPreClamp);
tonTurnLoss(IN := bTurnDriveInt AND (NOT rTrigTurn.Q), PT := tTurnLoss);
tonCutTo(IN := (eStateInt = E_DL_WrapSeqState.eCut) AND (NOT bCutDone), PT := tCutTimeout);
tonCutDwell(IN := NOT tonCutDwell.Q, PT := tCutDwell);
tonDwellHold(IN := (eStateInt = E_DL_WrapSeqState.eDwell), PT := tDwellHold);

(*------------------------------------------------------------------------------
 * 段 2｜上电首扫：计数与状态落安全侧
 *      First-scan init: counters and state to the safe side
 *-----------------------------------------------------------------------------*)
IF bFirstScan THEN
    eStateInt   := E_DL_WrapSeqState.eIdle;
    nBottomDone := 0;
    nTopDone    := 0;
    nRetryInt   := 0;
    bCutFailInt := FALSE;    // 首扫清切膜失败锁存 / Cut failure latch cleared on first scan
    bFirstScan  := FALSE;
END_IF

(*------------------------------------------------------------------------------
 * 段 3｜每拍预清（FB32-1）：单拍标志，禁入锁存 / 快照 / 计数
 *      Per-scan preset: single-scan flags only
 *-----------------------------------------------------------------------------*)
bErrorInt := FALSE;
bDoneT    := FALSE;

(*------------------------------------------------------------------------------
 * 段 4｜配方域闸（R151）+ 一致性核对：越界拒绝启动，不一致信息级按和执行
 *      Recipe gate and consistency check
 *      解除路径（R152 自证）：复位沿 AND 配方已改对
 *-----------------------------------------------------------------------------*)
bRecipeBad := (nBottomTurns < 1) OR (nBottomTurns > DL_WR_TURNS_MAX)
              OR (nTopTurns < 1) OR (nTopTurns > DL_WR_TURNS_MAX);

IF bRecipeBad THEN
    bRecipeLatch := TRUE;
    uErrorId     := 16#0005_03A9;    // 故障级：配方组态非法 / Fault: recipe illegal
    bErrorInt    := TRUE;
END_IF

bTotalDiff := (nTotalTurns <> (nBottomTurns + nTopTurns));
IF bTotalDiff AND (NOT bRecipeBad) THEN
    uErrorId := 16#0005_04D2;        // 信息级：总数不一致按和执行 / Info: total mismatch
END_IF

(*------------------------------------------------------------------------------
 * 段 5｜暂停双源合并与圈边界生效（ISA-88 相语义次源）
 *      Pause dual-source merge with turn-boundary effectiveness
 *      拍 N 进入：膜断 / 暂停请求置挂起；本拍行为：当前圈转完（沿到）即保持；
 *      拍 N+1 转出：请求撤销即恢复圈数继续（不重头）
 *-----------------------------------------------------------------------------*)
bPausePend := bFilmBreak OR bPauseReq;

IF fbTrigFilm.Q AND bPausePend THEN
    uErrorId := 16#0005_04D1;        // 信息级：膜断事件 / Info: film break event
END_IF

IF bPausePend AND rTrigTurn.Q THEN
    bPauseHoldInt := TRUE;           // 圈边界：暂停保持生效 / Boundary: pause hold engages
ELSIF NOT bPausePend THEN
    bPauseHoldInt := FALSE;          // 请求撤销：恢复 / Request gone: resume
END_IF

(*------------------------------------------------------------------------------
 * 段 6｜主状态机（红线 R6）：ENUM + CASE + ELSE 兜底
 *      Main state machine with the mandatory ELSE fallback
 *-----------------------------------------------------------------------------*)
CASE eStateInt OF

    E_DL_WrapSeqState.eIdle:
        (* eIdle 相执行输出清零（R57）：本相不写任何执行输出，出口段按状态归零 *)
        (* Idle clears outputs: the exit section derives all-off from the state *)
        (* 锁存驻留声明：反馈丢失 / 配方锁存的复位消化在 eFault 分支与空闲复位行处理 *)
        (* Latch dwell note: clears happen in the eFault branch and the idle reset line *)
        IF bReset THEN
            bTurnLossInt := FALSE;   // 空闲相复位也允许清反馈丢失锁存 / Idle reset clears loss latch
            bRecipeLatch := FALSE;   // 空闲相复位清配方锁存 / Idle reset clears recipe latch
            bCutFailInt  := FALSE;   // 空闲相复位清切膜失败锁存 / Idle reset clears cut failure latch
            uErrorId     := 16#0000_0000;
        END_IF
        IF bEnable AND (NOT bRecipeLatch) AND (NOT bTurnLossInt) AND (NOT bCutFailInt) AND fbTrigStart.Q THEN
            nBottomDone  := 0;       // 圈数计数清零 / Turn counters cleared
            nTopDone     := 0;
            nRetryInt    := 0;
            bPauseHoldInt := FALSE;
            eStateInt    := E_DL_WrapSeqState.ePreClamp;
        END_IF

    E_DL_WrapSeqState.ePreClamp:
        IF bStopCmd OR (NOT bEnable) THEN
            eStateInt := E_DL_WrapSeqState.eIdle;    // 退出 / Exit
        ELSIF bPreClampFb OR tonPre.Q THEN
            eStateInt := E_DL_WrapSeqState.eBottom;  // 反馈到位或建压窗满（双出口 R98）/ Feedback or window full
        END_IF

    E_DL_WrapSeqState.eBottom:
        IF bStopCmd OR (NOT bEnable) THEN
            eStateInt := E_DL_WrapSeqState.eIdle;
        ELSIF nBottomDone >= nBottomTurns THEN
            eStateInt := E_DL_WrapSeqState.eTop;     // 底圈数满转顶圈 / Bottom full, to top
        END_IF

    E_DL_WrapSeqState.eTop:
        IF bStopCmd OR (NOT bEnable) THEN
            eStateInt := E_DL_WrapSeqState.eIdle;
        ELSIF (nBottomDone + nTopDone) >= (nBottomTurns + nTopTurns) THEN
            eStateInt := E_DL_WrapSeqState.eCut;     // 总圈数满转切膜（验收：2+3=5）/ Total full, to cut
        END_IF

    E_DL_WrapSeqState.eCut:
        IF bStopCmd OR (NOT bEnable) THEN
            eStateInt := E_DL_WrapSeqState.eIdle;
        ELSIF bCutDone THEN
            eStateInt := E_DL_WrapSeqState.eDwell;   // 切膜完成进保持 / Cut done, to dwell
        END_IF

    E_DL_WrapSeqState.eDwell:
        IF bStopCmd OR (NOT bEnable) THEN
            eStateInt := E_DL_WrapSeqState.eIdle;
        ELSIF tonDwellHold.Q THEN
            bDoneT    := TRUE;       // 完成脉冲：内部置位 -> 出口单拍映射（两段式）/ Done pulse via exit
            eStateInt := E_DL_WrapSeqState.eIdle;
        END_IF

    E_DL_WrapSeqState.eFault:
        (* 解除路径（R152 自证可达）：复位沿 AND 反馈已恢复 AND 配方已改对 *)
        (* 三类锁存同沿解除：配方 / 反馈丢失 / 切膜失败（人工复位是切膜失败的唯一出路） *)
        IF fbTrigReset.Q AND (NOT bRecipeBad) THEN
            bRecipeLatch := FALSE;
            bTurnLossInt := FALSE;
            bCutFailInt  := FALSE;       // 切膜失败锁存解除（人工复位）/ Cut failure latch cleared by the manual reset
            uErrorId     := 16#0000_0000;
            eStateInt    := E_DL_WrapSeqState.eIdle;
        END_IF

    ELSE
        (* 非法状态拦截：迁兜底态（复用配方段码位） *)
        eStateInt := E_DL_WrapSeqState.eFault;
        uErrorId  := 16#0005_03A9;
        bErrorInt := TRUE;

END_CASE;

(*------------------------------------------------------------------------------
 * 段 7｜转盘圈计数（沿计数 + 饱和 255）与反馈丢失消化
 *      Turn counting with 255 saturation, and the feedback loss digestion
 *      计数仅在驱动输出有效且未暂停保持时推进（暂停在圈边界已截停驱动）
 *-----------------------------------------------------------------------------*)
bTurnDriveInt := (eStateInt = E_DL_WrapSeqState.eBottom) OR (eStateInt = E_DL_WrapSeqState.eTop);
bTurnDriveInt := bTurnDriveInt AND (NOT bPauseHoldInt);

IF rTrigTurn.Q AND bTurnDriveInt THEN
    (* 终审就地修 v1.0.1（R68④）：计数上限改用总圈上界 510。原实现以单段上界 255
     * 作总数闸，配方合法（如底 200 + 顶 100 = 300）时计数停在 255 -> eTop 相
     * 永不可达、转盘驱动常励磁（死路径）。 *)
    (* The counter ceiling is the total bound, so legal recipes above 255 turns no longer deadlock. *)
    IF (nBottomDone + nTopDone) < DL_WR_TOTAL_MAX THEN
        IF eStateInt = E_DL_WrapSeqState.eBottom THEN
            nBottomDone := nBottomDone + 1;  // 底圈计数推进 / Bottom count up
        ELSIF eStateInt = E_DL_WrapSeqState.eTop THEN
            nTopDone := nTopDone + 1;        // 顶圈计数推进 / Top count up
        END_IF
    END_IF
END_IF

IF tonTurnLoss.Q AND (NOT bTurnLossInt) THEN
    bTurnLossInt := TRUE;            // 反馈丢失锁存 / Loss latched
    uErrorId     := 16#0005_03AA;    // 故障级：反馈丢失 / Fault: feedback loss
    bErrorInt    := TRUE;
    eStateInt    := E_DL_WrapSeqState.eFault;   // 锁存同步迁相（FB50-1④）/ Latch migrates phase
END_IF

(*------------------------------------------------------------------------------
 * 段 8｜切膜重试节流、计数饱和与失败出口（R69 点修②）
 *      Film cut retry throttle, count saturation and the failure exit
 *      重试由自复位间隔窗节流：每窗到期 +1 次（防同拍连发）；
 *      计次饱和（nCutRetryMax 封顶不回绕）后**不再自动重切**：单次窗再次超时即判
 *      切膜失败 -> 03B3 + bCutFail 锁存 + 迁 eFault 停机待人工，解除靠人工复位。
 *      nCutRetryMax <= 0 表示「不允许重试」，首次窗超时即判失败（安全侧直落）。
 *-----------------------------------------------------------------------------*)
IF (eStateInt = E_DL_WrapSeqState.eCut) AND tonCutTo.Q THEN
    IF nRetryInt >= nCutRetryMax THEN
        (* 拍 N 进入：计次已饱和且单次窗再次超时；本拍行为：锁存失败码并迁故障相，
         * 拒绝任何自动重切；拍 N+1 转出：eFault 驻留至人工复位沿。 *)
        (* Retries exhausted and the cut window expired again: latch the failure, never retry automatically *)
        bCutFailInt := TRUE;         // 切膜失败锁存 / Cut failure latched
        uErrorId    := 16#0005_03B3; // 故障级：切膜失败，停机待人工 / Fault: cut failed, manual service
        bErrorInt   := TRUE;         // R45 配对 / Paired with the fault code
        eStateInt   := E_DL_WrapSeqState.eFault;   // 锁存同步迁相 / Latch migrates phase
    ELSIF tonCutDwell.Q THEN
        (* 双窗合流节流：切膜窗保持超时的同时，重试间隔窗到期才计一次（防同拍连发） *)
        (* Double-window throttle: count at most once per dwell period while timed out *)
        IF nRetryInt < nCutRetryMax THEN
            nRetryInt := nRetryInt + 1;  // 重试计数推进 / Retry count up
        END_IF
        IF nRetryInt >= nCutRetryMax THEN
            uErrorId := 16#0005_04D3;    // 信息级：重试已饱和，下一窗超时即判失败 / Info: retries saturated
        END_IF
    END_IF
END_IF

(*------------------------------------------------------------------------------
 * 段 9｜输出单一出口（范式 P-05）
 *      Single output exit
 *-----------------------------------------------------------------------------*)
bTurnDrive   := bTurnDriveInt AND (NOT bTurnLossInt) AND (NOT bCutFailInt);
(* 压膜出口（R69 点修⑦）：仅 ePreClamp 相有效；底 / 顶圈段一进入即释放并全程保持
 * 释放（防膜皱 / 拉断），切膜 / 保持 / 空闲 / 故障相同样释放。释放由状态派生式
 * 结构性保证，不挂单拍标志，也不受暂停位改写。 *)
(* Press-film output is only driven in the pre-clamp phase; the winding phases stay released *)
bPreClampOut := (eStateInt = E_DL_WrapSeqState.ePreClamp);
bCutOut      := (eStateInt = E_DL_WrapSeqState.eCut) AND (NOT bCutDone) AND (NOT bCutFailInt);
bCutFail     := bCutFailInt;         // 失败锁存直出（人工复位前常驻）/ Failure latch straight out
bPauseHold   := bPauseHoldInt;
bSeqActive   := (eStateInt <> E_DL_WrapSeqState.eIdle) AND (eStateInt <> E_DL_WrapSeqState.eFault);
bSeqDone     := bDoneT;              // 完成脉冲统一出口（预清 + 两段式）/ Unified done exit
nTurnsDone   := nBottomDone + nTopDone;
nCutRetries  := nRetryInt;
bError       := bErrorInt OR (eStateInt = E_DL_WrapSeqState.eFault);
eState       := eStateInt;
END_FUNCTION_BLOCK

(* ---- FB_DL_StringFifoRetry.st ---- *)
(*==============================================================================
 * 组件名称 (Component)  : FB_DL_StringFifoRetry
 * 所属子库 (Sublibrary) : DL_Process
 * 当前版本 (Version)    : 1.0.0
 * 兼容性   (Platform)   : CODESYS 3.5+ / TwinCAT 3 / 汇川 InoProShop / 施耐德 Machine Expert
 *                         仅依赖 Standard.library（TON / R_TRIG / LEN），零厂商私有库
 * 功能描述 (Function)   : 电池串缓存队列重试出站。
 *                         上游把电池串编号压入定长缓冲，本件按 FIFO 逐条向 MES/贴标工位出站，
 *                         每条出站走"发令 → 等确认 → 成功出队 / 失败计数"的握手闭环；
 *                         同一串失败重试超上限即锁存 NG 并停线等人工复位。
 *                         三条固化纪律：
 *                           ① **丢新策略**：队满时丢弃**新到**的串、保留已在队旧串
 *                              （旧串已在产线中途，丢旧会切断履历；丢新只丢一条未开始处理的串）；
 *                           ② **重试计数上限**：nMaxRetries 提为引脚（禁魔法数），
 *                              达到上限即锁存 bRetryNg；上限域闸 nMaxRetries ≥ 1；
 *                           ③ **单拍脉冲两段式**：发令脉冲 _bTxValid 在 CASE 内用内部位
 *                              置位、段 8 统一映射出口，禁同相内置位后同相撤位（R129）。
 *                         验收向量：
 *                           ① 深度 16；压入 16 条后续压 → 丢新 + eDroppedNew（信息级，不锁存）
 *                           ② nMaxRetries = 3；同一条连续 3 次 bAckFail → 第 3 次锁存 bRetryNg
 *                           ③ 握手超时 tHandshakeTo 到 → 计一次失败（与 bAckFail 同权）
 *                           ④ bAckOk 到达 → 出队、重试计数清零、回 eIdle
 * 接口     (Interface)  : 入 bPush 入队沿、sInString 入队电池串、bStart 出站使能、bAckOk 下游确认、
 *                         bAckFail 下游失败、nMaxRetries 重试上限、tHandshakeTo 握手超时、
 *                         bReset 复位沿；
 *                         出 sTxString 当前出站串、bTxValid 发令脉冲（单拍）、bTxBusy 等确认中、
 *                         iRetryCnt 当前串已试次数、iQueueCnt 在队条数、bDropped 当拍丢新、
 *                         bRetryNg 重试超限锁存、eState 相、eCause 成因、bError 故障标志。
 * 边界     (Boundary)   : ① **属主边界（写死）：本件只管"缓冲区与重试编排"，不做报文编码/
 *                         串口收发/协议校验**（属通讯层件），也不判电池串数据内容是否合法；
 *                         ② **深度闸**：环形指针与槽位下标一律钳在 1..16（字面量上界），
 *                         同值常量 DL_SFR_DEPTH 作运行时二次闸（R104）；
 *                         ③ **超时监视冻结**：tonHandshake 的 IN 串 (NOT _bFault)，
 *                         故障期间不累计，复位同拍不会立即重锁（R252 第 2 变体）；
 *                         ④ **重试上限域闸**：nMaxRetries ≤ 0 → 锁存 eCfgIllegal（零上限会让
 *                         第 0 次即判超限，属静默失效 R179）；
 *                         ⑤ **锁存解除式**：bRetryNg / eFault 的解除仅 bReset 上升沿
 *                         （R228B 唯一迁出）；bReset 为外部引脚，不受锁存量门控，恒可达；
 *                         ⑥ 零全局耦合、零物理地址。
 * 分工声明 (Scope)      : 本件只管"电池串缓存队列的出站重试"。不接管：底层 FIFO 结构件
 *                         （FB_DL_FifoBuffer 族）、MES 报文重传的幂等去重（属通讯层）、
 *                         电池串工艺合格判定（属测试判据件）。
 * 来源标签 (Source Tag) : ROADMAP 空勾真缺口 P1（电池串重试出站，自研 clean-room）
 * 码表     (Codes)      : 本件不占用任何全局数字码位（零码位范式 R297）；诊断由 BOOL + ENUM 出口承担。
 * 红线自检 (Redline)    : R1 ✓ 零 GVL/VAR_EXTERNAL ｜ R2 ✓ 零 %I/%Q/%M ｜ R3 ✓ 纯 IEC 61131-3
 *                         R4 ✓ 指针钳位 + 上限域闸 + 重试计数饱和 ｜ R5 ✓ 声明逐行同行双语注释
 *                         R6 ✓ ENUM+CASE 含 ELSE 兜底 ｜ R7 ✓ TON/四 R_TRIG 段 0 无条件刷新
 * 修订历史 (Revision)   : 2026-11-19  v1.0.0  R47 首版（批次 2 · 序号 7）
 *==============================================================================*)

TYPE E_DL_SfrState :
(
    eIdle    := 0,    // 待机相（可取队首出站） / Idle, ready to take the head record
    eWaitAck := 10,   // 等确认相（握手窗口内） / Waiting for the downstream acknowledgement
    eFault   := 90    // 故障相（等复位） / Fault, awaiting reset
);
END_TYPE

TYPE E_DL_SfrCause :
(
    eNone        := 0,   // 无异常 / No anomaly
    eCfgIllegal  := 1,   // 组态非法（重试上限非正） / Illegal configuration, retry limit non-positive
    eDroppedNew  := 2,   // 队满丢新（信息级） / Queue full, newest dropped, info level
    eStringEmpty := 3,   // 入队空串（信息级） / Empty string rejected, info level
    eAckFail     := 4,   // 下游失败（计数未超限，信息级） / Downstream failure below the retry limit
    eHsTimeout   := 5,   // 握手超时（计数未超限，信息级） / Handshake timeout below the retry limit
    eRetryNg     := 6,   // 重试超限（锁存，故障级） / Retry limit exceeded, latched
    ePtrCorrupt  := 7,   // 环形指针损坏（故障级） / Ring pointer corruption, fault level
    ePhaseBad    := 8    // 非法相位兜底 / Illegal phase fallback
);
END_TYPE

FUNCTION_BLOCK FB_DL_StringFifoRetry
VAR_INPUT
    bPush        : BOOL := FALSE;       // 入队沿 [-] / Enqueue edge
    sInString    : STRING[63] := '';    // 待入队电池串编号 [-] / Cell-string identifier to enqueue
    bStart       : BOOL := FALSE;       // 出站使能（TRUE 时自动取队首出站） [-] / Outbound enable
    bAckOk       : BOOL := FALSE;       // 下游确认成功（当拍电平） [-] / Downstream acknowledgement, level
    bAckFail     : BOOL := FALSE;       // 下游失败（当拍电平） [-] / Downstream failure, level
    nMaxRetries  : INT := 3;            // 单串重试上限，域 ≥ 1 [次] / Retry limit per string, domain >= 1
    tHandshakeTo : TIME := T#3S;        // 握手超时，域 > T#0S [ms] / Handshake timeout, > T#0S [ms]
    bReset       : BOOL := FALSE;       // 复位沿（清故障锁存与重试计数） [-] / Reset edge
END_VAR
VAR_OUTPUT
    sTxString : STRING[63] := '';                        // 当前出站电池串 [-] / String currently being transmitted
    bTxValid  : BOOL := FALSE;                           // 发令脉冲（单拍） [-] / Transmit pulse, single scan
    bTxBusy   : BOOL := FALSE;                           // 等确认中 [-] / Waiting for acknowledgement
    iRetryCnt : INT := 0;                                // 当前串累计失败次数 [次] / Failure count of the current string
    iQueueCnt : INT := 0;                                // 在队条数 [条] / Records currently queued
    bDropped  : BOOL := FALSE;                           // 当拍发生丢新 [-] / Newest record dropped this scan
    bRetryNg  : BOOL := FALSE;                           // 重试超限锁存（等复位） [-] / Retry limit exceeded, latched
    eState    : E_DL_SfrState := E_DL_SfrState.eIdle;    // 相出口 [-] / Phase outlet
    eCause    : E_DL_SfrCause := E_DL_SfrCause.eNone;    // 成因出口（R190 归因唯一） [-] / Cause outlet
    bError    : BOOL := FALSE;                           // 故障标志（仅故障级成因） [-] / Error flag, fault level only
END_VAR
VAR
    _eState    : E_DL_SfrState := E_DL_SfrState.eIdle;   // 内部相（CASE 唯一写入目标） / Internal phase
    _eCause    : E_DL_SfrCause := E_DL_SfrCause.eNone;   // 成因锁存量 / Latched cause
    _bFault    : BOOL := FALSE;                          // 故障锁存位 / Latched fault bit
    _bRetryNg  : BOOL := FALSE;                          // 重试超限锁存位 / Latched retry-NG bit
    _iHead     : INT := 1;                               // 队列头指针（1..16） / Queue head pointer
    _iTail     : INT := 1;                               // 队列尾指针（1..16） / Queue tail pointer
    _iCnt      : INT := 0;                               // 在队条数 / Queued count
    _iRetry    : INT := 0;                               // 当前串失败计数 / Failure count of the current string
    _sTx       : STRING[63] := '';                       // 当前出站串内部副本 / Internal copy of the transmitting string
    _bTxValid  : BOOL := FALSE;                          // 发令脉冲内部位（单拍） / Internal transmit pulse
    _bDropped  : BOOL := FALSE;                          // 丢新内部位（单拍） / Internal drop flag
    _bCfgBad   : BOOL := FALSE;                          // 组态非法当拍量 / Illegal configuration this scan
    _bConsume  : BOOL := FALSE;                          // 本拍应消费队首（成功出队） / Head should be consumed this scan
    _bFailArmed: BOOL := TRUE;                           // 失败条件武装位（沿消费一次，条件消失后重武装） / Failure-edge arming flag
    tonHs      : TON;                                    // 握手超时实例，段 0 无条件调用 / Handshake timeout instance
    rtPush     : R_TRIG;                                 // 入队沿实例，段 0 无条件调用 / Enqueue edge instance
    rtReset    : R_TRIG;                                 // 复位沿实例，段 0 无条件调用 / Reset edge instance
    asBuf      : ARRAY[1..16] OF STRING[63];             // 电池串环（深度字面量上界，R104） / String ring, literal depth
END_VAR
VAR CONSTANT
    DL_SFR_DEPTH : INT := 16;            // 队列深度（与数组字面量上界同源） [条] / Queue depth
    DL_SFR_RTY_MAX : INT := 100;         // 重试上限的工程上限保护 [次] / Engineering upper bound of the retry limit
END_VAR

(* —— 段 0：组态闸 + TON 与两沿无条件周期刷新（R228A；IN 串故障否决，R252） —— *)
_bCfgBad := (nMaxRetries <= 0) OR (nMaxRetries > DL_SFR_RTY_MAX) OR (tHandshakeTo <= T#0S);   // 上限须 1..100 且超时须为正
rtPush(CLK := bPush);                                    // 入队沿 / Enqueue edge
rtReset(CLK := bReset);                                  // 复位沿 / Reset edge
tonHs(IN := (_eState = E_DL_SfrState.eWaitAck) AND (NOT _bFault), PT := tHandshakeTo);   // 握手超时（等确认相派生） / Handshake timeout

(* —— 段 1：单拍量预清零（锁存量 _eCause/_bFault/_bRetryNg/_iRetry 不入清单，R107） —— *)
_bTxValid := FALSE;                                      // 发令脉冲预清 / Transmit pulse preset
_bDropped := FALSE;                                      // 丢新标志预清 / Drop flag preset
bError    := FALSE;                                      // 故障标志预清（R45 配对） / Error preset

(* —— 段 2：组态闸（非法即锁存故障级） —— *)
IF _bCfgBad THEN
    _eCause := E_DL_SfrCause.eCfgIllegal;                // 归因：组态非法 / Cause: illegal configuration
    _bFault := TRUE;                                     // 锁存 / Latch
    _eState := E_DL_SfrState.eFault;                     // 入故障相 / Enter fault phase
END_IF

(* —— 段 3：环形指针自检（越界即清队重建 + 锁存） —— *)
IF (_iHead < 1) OR (_iHead > DL_SFR_DEPTH) OR (_iTail < 1) OR (_iTail > DL_SFR_DEPTH)
   OR (_iCnt < 0) OR (_iCnt > DL_SFR_DEPTH) THEN
    _iHead := 1;                                         // 头指针重建 / Head rebuilt
    _iTail := 1;                                         // 尾指针重建 / Tail rebuilt
    _iCnt  := 0;                                         // 计数清零 / Count cleared
    _eCause := E_DL_SfrCause.ePtrCorrupt;                // 归因：指针损坏 / Cause: pointer corruption
    _bFault := TRUE;                                     // 锁存 / Latch
    _eState := E_DL_SfrState.eFault;                     // 入故障相 / Enter fault phase
END_IF

(* —— 段 4：迁出链（bReset 唯一迁出：清故障锁存 + 重试计数 + 相位；R228B） —— *)
IF rtReset.Q THEN
    _bFault   := FALSE;                                  // 清故障锁存 / Clear fault latch
    _bRetryNg := FALSE;                                  // 清重试超限锁存 / Clear retry-NG latch
    _eCause   := E_DL_SfrCause.eNone;                    // 清成因 / Clear cause
    _iRetry   := 0;                                      // 重试计数清零 / Retry counter cleared
    _iHead    := 1;                                      // 头指针回 1（队列随之作废） / Head back to 1, queue discarded
    _iTail    := 1;                                      // 尾指针回 1 / Tail back to 1
    _iCnt     := 0;                                      // 计数清零 / Count cleared
    _sTx      := '';                                     // 出站副本清空 / Transmit copy cleared
    _eState   := E_DL_SfrState.eIdle;                    // 回待机相 / Back to idle
END_IF

(* —— 段 5：入队（丢新策略：满则丢新、保旧；空串拒入） —— *)
IF (rtPush.Q) AND (NOT _bFault) THEN
    IF LEN(sInString) = 0 THEN
        _eCause := E_DL_SfrCause.eStringEmpty;           // 归因：空串拒入（信息级） / Cause: empty string, info level
    ELSIF _iCnt >= DL_SFR_DEPTH THEN
        _bDropped := TRUE;                               // 丢新锁存（当拍） / Drop the newest record
        _eCause := E_DL_SfrCause.eDroppedNew;            // 归因：队满丢新（信息级） / Cause: full, newest dropped
    ELSE
        asBuf[_iTail] := sInString;                      // 写尾槽位 / Write the tail slot
        _iCnt  := _iCnt + 1;                             // 计数递增 / Count increment
        _iTail := _iTail + 1;                            // 尾指针推进 / Tail advance
        IF _iTail > DL_SFR_DEPTH THEN
            _iTail := 1;                                 // 环形回卷 / Ring wrap
        END_IF
    END_IF
END_IF

(* —— 段 6：相迁移（出站握手闭环） —— *)
IF (NOT _bFault) AND (NOT _bCfgBad) THEN
    CASE _eState OF

    E_DL_SfrState.eIdle:
        IF bStart AND (_iCnt > 0) THEN
            _sTx      := asBuf[_iHead];                  // 取队首出站串 / Take the head string
            _bTxValid := TRUE;                           // 发令脉冲（内部位，段 8 单点映射） / Internal transmit pulse
            _iRetry   := 0;                              // 新串重试计数归零 / Reset the retry counter for the new string
            _eState   := E_DL_SfrState.eWaitAck;         // 进等确认相 / Enter the wait-ack phase
        END_IF

    E_DL_SfrState.eWaitAck:
        IF bAckOk THEN
            _bConsume := TRUE;                           // 成功：本拍消费队首 / Success: consume the head this scan
            _iRetry   := 0;                              // 重试计数归零 / Retry counter cleared
            _eState   := E_DL_SfrState.eIdle;            // 回待机相 / Back to idle
        ELSIF (bAckFail OR tonHs.Q) AND _bFailArmed THEN
            _bFailArmed := FALSE;                        // 失败条件沿消费一次（条件消失后重新武装，防每拍累加） / Consume the failure edge once
            _iRetry := _iRetry + 1;                      // 失败计数 +1（失败与超时同权） / Failure or timeout, same weight
            IF bAckFail THEN
                _eCause := E_DL_SfrCause.eAckFail;       // 归因：下游失败 / Cause: downstream failure
            ELSE
                _eCause := E_DL_SfrCause.eHsTimeout;     // 归因：握手超时 / Cause: handshake timeout
            END_IF
            IF _iRetry >= nMaxRetries THEN
                _bRetryNg := TRUE;                       // 重试超限锁存 / Latch the retry-NG state
                _bFault   := TRUE;                       // 故障锁存 / Latch the fault
                _eCause   := E_DL_SfrCause.eRetryNg;     // 归因：重试超限（覆盖为故障级首因） / Cause: retry limit, fault level
                _eState   := E_DL_SfrState.eFault;       // 入故障相（等复位） / Enter the fault phase
            ELSE
                _bTxValid := TRUE;                       // 未超限：当拍重发（内部位） / Below the limit: retransmit
                _eState   := E_DL_SfrState.eWaitAck;     // 留在等确认相 / Stay in the wait-ack phase
            END_IF
        END_IF

    E_DL_SfrState.eFault:
        ;                                            // 故障相：仅等复位沿 / Wait for the reset edge only

    ELSE
        _eCause := E_DL_SfrCause.ePhaseBad;              // 归因：非法相位 / Cause: illegal phase
        _bFault := TRUE;                                 // 锁存 / Latch
        _eState := E_DL_SfrState.eFault;                 // 强拉故障相 / Force fault phase

    END_CASE
END_IF

(* —— 段 6b：失败条件消失后重新武装（沿消费纪律；锁存量不入每拍预清零） —— *)
IF (NOT bAckFail) AND (NOT tonHs.Q) THEN
    _bFailArmed := TRUE;                                 // 条件消失：重新武装 / Condition gone: re-arm
END_IF

(* —— 段 7：出队（成功消费唯一入口；指针回卷） —— *)
IF _bConsume THEN
    asBuf[_iHead] := '';                                 // 清空已发送槽位 / Clear the sent slot
    _iCnt  := _iCnt - 1;                                 // 计数递减 / Count decrement
    _iHead := _iHead + 1;                                // 头指针推进 / Head advance
    IF _iHead > DL_SFR_DEPTH THEN
        _iHead := 1;                                     // 环形回卷 / Ring wrap
    END_IF
    _bConsume := FALSE;                                  // 消费标志自复位（防跨拍误消费） / Self-reset the consume flag
END_IF

(* —— 段 8：出口单点映射（名实双出口，R191） —— *)
sTxString := _sTx;                                       // 当前出站串出口 / Transmit string outlet
bTxValid  := _bTxValid;                                  // 发令脉冲出口 / Transmit pulse outlet
bTxBusy   := (_eState = E_DL_SfrState.eWaitAck);         // 等确认中出口 / Busy outlet
iRetryCnt := _iRetry;                                    // 失败计数出口 / Retry count outlet
iQueueCnt := _iCnt;                                      // 在队条数出口 / Queued count outlet
bDropped  := _bDropped;                                  // 丢新出口 / Drop outlet
bRetryNg  := _bRetryNg;                                  // 重试超限出口 / Retry-NG outlet
eState    := _eState;                                    // 相出口 / Phase outlet
eCause    := _eCause;                                    // 成因出口 / Cause outlet
bError    := _bFault;                                    // 故障标志 / Error flag

END_FUNCTION_BLOCK

(* ---- FB_DL_TabWeldingMonitor.st ---- *)
(*==============================================================================
 * 组件名称 (Component)  : FB_DL_TabWeldingMonitor
 * 所属子库 (Sublibrary) : DL_Process
 * 当前版本 (Version)    : 1.0.1
 * 兼容性   (Platform)   : CODESYS 3.5+ / TwinCAT 3 / 汇川 InoProShop / 施耐德 Machine Expert
 *                         仅依赖 Standard.library（R_TRIG），零厂商私有库
 * 功能描述 (Function)   : 极耳焊能量/位移/压力三包络窗口判定。每次焊接结束时由 bEval 上升沿触发
 *                         一次评估，在**同一拍内**对三路各判一次双侧包络（下限与上限都要查，
 *                         只查上限会漏"欠能量虚焊"这类最常见的失效）：
 *                           能量 fEnergy ∈ [fEnergyLo, fEnergyHi]  → 否则 bEnergyNg
 *                           位移 fDisp   ∈ [fDispLo,   fDispHi]    → 否则 bDispNg
 *                           压力 fPressure ∈ [fPressLo, fPressHi]  → 否则 bPressNg
 *                         三路**独立**判定、**独立**故障位，绝不合并成一个"焊接不良"位：
 *                         合并后无法区分是能量不足还是压力不足，工艺调参无从下手。
 *                         另出 nNgMask 通道位掩码（bit0 能量 / bit1 位移 / bit2 压力）便于 HMI
 *                         一字节展示，但台账判定仍以三个 BOOL 为准（掩码是展示便利，不是判据）。
 *                         任一通道越窗 → bAnyNg 锁存（累计），直到 bReset 上升沿才清，
 *                         保证两次评估之间的 NG 不会被下一次合格件抹掉（R187 锁存纪律）。
 * 接口     (Interface)  : 输入 fEnergy / fDisp / fPressure 三路实测、六个包络阈值、bEval 评估沿、
 *                         bReset 复位；输出 bEnergyNg / bDispNg / bPressNg 三路独立故障位（锁存）、
 *                         bAnyNg 任一路故障（锁存）、nNgMask 通道位掩码、bEvalDone 单拍评估完成、
 *                         eState / eCause / bError。
 * 边界     (Boundary)   : ① **属主边界（写死）：本件只做"一次焊点的三包络判定"，不控制焊接电源、
 *                         不排序焊点、不判焊点位置**。焊接时序与焊点序列属焊接主控 POU；
 *                         本件的结论位供主控做 NG 剔除与工艺趋势。
 *                         ② 组态闸（每个参与判据的引脚都要闸，缺一即该通道恒判 NG 或恒判 OK）：
 *                         六条阈值任一 fXxxLo >= fXxxHi（上下限倒置）、任一引脚 NaN → 故障锁存，
 *                         三个通道同时不宣称结果（bEvalDone 不出，避免把闸门故障记成焊点 NG）。
 *                         ③ 评估是"沿触发单拍"语义：非评估拍不改变任何锁存位，也不清位。
 *                         ④ 单枚 R_TRIG（bEval）与单枚 R_TRIG（bReset）段 0 无条件周期刷新；
 *                         本件无 TON，故无跨相复位风险。
 *                         ⑤ 故障相迁出唯一路径 = bReset 上升沿（R228B）。
 *                         ⑥ 零全局耦合（无 GVL / 无 VAR_EXTERNAL / 无物理地址）。
 * 分工声明 (Scope)      : 与 `FB_DL_AxisTorqueLimitGuard`（轴力矩瞬时限）分工——那件在运动中连续
 *                         判力矩，本件在焊后一次性判三包络；时间语义（连续 vs 单点）不同，不可互替。
 * 来源标签 (Source Tag) : ROADMAP B 类（锂电池极耳焊工艺监控，自研 clean-room，无外源代码）
 * 解除式   (Release)    : bReset 上升沿 ∧ 组态合法 → 清三路 NG 与任一路 NG 锁存。
 *                         自证可满足：复位为外部动作，不受判据门控；清后下一评估沿重新判定。
 * 码表     (Codes)      : 本件不占用任何全局数字码位。故障出口为三个独立 BOOL + BYTE 通道掩码
 *                         （掩码是**通道位**，不是全局事件码，不参与码段分配）；数字码位待主控
 *                         收口阶段统一派号。
 * 红线自检 (Redline)    : R1 ✓ 零 GVL/VAR_EXTERNAL ｜ R2 ✓ 零 %I/%Q/%M ｜ R3 ✓ 纯 IEC 61131-3
 *                         R4 ✓ 六阈值双侧几何闸 + NaN 闸 + 浮点容差 ｜ R5 ✓ 声明逐行同行双语注释
 *                         R6 ✓ ENUM+CASE 含 ELSE ｜ R7 ✓ R_TRIG 段 0 无条件刷新
 * 返修记录 (Repair)     : v1.0.1（R47 P0 返修）实测 NaN 单列 eMeasBad 出口：原先实测与阈值非有限并入同一
 *                         eCfgIllegal 并锁存，传感器瞬时掉线会把 HMI 打到"组态非法"（误导维护方向）。
 *                         现改为——实测类 NaN 当拍跳过评估、只置 eMeasBad、不锁存、不动通道位；
 *                         阈值类 NaN 与阈值倒置仍判 eCfgIllegal 并锁存（须人工修参数）。
 * 修订历史 (Revision)   : 2026-11-19  v1.0.0  R46 首版（批次 2 · 序号 10）
 *==============================================================================*)

TYPE E_DL_TwmState :
(
    eIdle  := 0,    // 等待首次评估沿 / Awaiting the first evaluation edge
    eRun   := 10,   // 逐焊点评估运行相 / Evaluating per weld spot
    eFault := 90    // 组态故障相 / Configuration fault phase
);
END_TYPE

TYPE E_DL_TwmCause :
(
    eNone       := 0,   // 无异常 / No anomaly
    eCfgIllegal := 1,   // 组态非法（阈值倒置或非有限） / Illegal configuration
    eEnergyNg   := 2,   // 能量越窗 / Energy out of the envelope
    eDispNg     := 3,   // 位移越窗 / Displacement out of the envelope
    ePressNg    := 4,   // 压力越窗 / Pressure out of the envelope
    eMultiNg    := 5,   // 多路同时越窗（归因无法唯一，单列成因） / Multiple channels out of the envelope
    eMeasBad    := 6,   // 实测值 NaN（当拍跳过评估，不锁存） / Measured value NaN, scan skipped, not latched
    ePhaseBad   := 7    // 非法相位兜底 / Illegal phase fallback
);
END_TYPE

FUNCTION_BLOCK FB_DL_TabWeldingMonitor
VAR_INPUT
    fEnergy   : REAL := 0.0;     // 焊接能量实测 [J] / Measured weld energy [J]
    fDisp     : REAL := 0.0;     // 焊接位移实测（电极下压量） [mm] / Measured displacement [mm]
    fPressure : REAL := 0.0;     // 焊接压力实测 [N] / Measured weld pressure [N]
    fEnergyLo : REAL := 10.0;    // 能量窗下限，域 < fEnergyHi [J] / Energy lower envelope, < upper [J]
    fEnergyHi : REAL := 100.0;   // 能量窗上限，域 > fEnergyLo [J] / Energy upper envelope, > lower [J]
    fDispLo   : REAL := 0.05;    // 位移窗下限，域 < fDispHi [mm] / Displacement lower envelope [mm]
    fDispHi   : REAL := 1.50;    // 位移窗上限，域 > fDispLo [mm] / Displacement upper envelope [mm]
    fPressLo  : REAL := 50.0;    // 压力窗下限，域 < fPressHi [N] / Pressure lower envelope [N]
    fPressHi  : REAL := 500.0;   // 压力窗上限，域 > fPressLo [N] / Pressure upper envelope [N]
    bEval     : BOOL := FALSE;   // 评估触发，上升沿判一次 [-] / Evaluation trigger, judges once per rising edge
    bReset    : BOOL := FALSE;   // 复位，上升沿清三路 NG 锁存 [-] / Reset, rising edge clears NG latches
END_VAR
VAR_OUTPUT
    bEnergyNg : BOOL;               // 能量越窗（锁存） [-] / Energy out of envelope, latched
    bDispNg   : BOOL;               // 位移越窗（锁存） [-] / Displacement out of envelope, latched
    bPressNg  : BOOL;               // 压力越窗（锁存） [-] / Pressure out of envelope, latched
    bAnyNg    : BOOL;               // 任一路越窗（锁存累计） [-] / Any channel out of envelope, latched
    nNgMask   : BYTE;               // 通道位掩码：bit0 能量 / bit1 位移 / bit2 压力 [-] / Channel bit mask, bit0 energy, bit1 displacement, bit2 pressure
    bEvalDone : BOOL;               // 本次评估完成，单拍脉冲 [-] / Evaluation completed, single-scan pulse
    eState    : E_DL_TwmState;      // 状态出口 [-] / State outlet
    eCause    : E_DL_TwmCause;      // 成因出口（R190 归因唯一） [-] / Cause outlet
    bError    : BOOL;               // 故障标志（组态故障或任一路 NG） [-] / Error flag
END_VAR
VAR
    _eState   : E_DL_TwmState := E_DL_TwmState.eIdle;    // 内部相位（CASE 唯一写入目标） / Internal phase
    _eCause   : E_DL_TwmCause := E_DL_TwmCause.eNone;    // 成因锁存量 / Latched cause
    rtEval    : R_TRIG;         // 评估沿实例，段 0 无条件调用 / Evaluation edge instance
    rtReset   : R_TRIG;         // 复位沿实例，段 0 无条件调用 / Reset edge instance
    _bNg1     : BOOL;           // 能量越窗锁存位（锁存量） / Latched energy NG
    _bNg2     : BOOL;           // 位移越窗锁存位（锁存量） / Latched displacement NG
    _bNg3     : BOOL;           // 压力越窗锁存位（锁存量） / Latched pressure NG
    _bAnyNg   : BOOL;           // 任一路越窗锁存位（锁存量） / Latched any-NG
    _bCfgBad  : BOOL;           // 组态非法当拍量 [-] / Illegal configuration this scan
    _bNonFin  : BOOL;           // 输入非有限当拍量（含阈值） [-] / Non-finite input this scan
    _bThBad   : BOOL;           // 阈值类非法当拍量（NaN 或倒置，锁存级） [-] / Threshold invalid, latched
    _bMeasBad : BOOL;           // 实测类 NaN 当拍量（跳过评估，不锁存） [-] / Measured NaN, skipped, not latched
    _bE1      : BOOL;           // 本次评估能量越窗当拍量 [-] / Energy NG this evaluation
    _bE2      : BOOL;           // 本次评估位移越窗当拍量 [-] / Displacement NG this evaluation
    _bE3      : BOOL;           // 本次评估压力越窗当拍量 [-] / Pressure NG this evaluation
    _nNgCnt   : USINT;          // 本次评估越窗通道计数（归因唯一性判据） [路] / Channels out of envelope this evaluation
END_VAR
VAR CONSTANT
    DL_TWM_MASK_E : BYTE := 16#01;   // 通道位掩码：能量 [位] / Channel mask bit for energy
    DL_TWM_MASK_D : BYTE := 16#02;   // 通道位掩码：位移 [位] / Channel mask bit for displacement
    DL_TWM_MASK_P : BYTE := 16#04;   // 通道位掩码：压力 [位] / Channel mask bit for pressure
END_VAR

(* —— 段 0：判据派生 + 两沿实例无条件周期刷新 —— *)
(* v1.0.1：实测 NaN 与阈值 NaN 分列——实测类当拍跳过不锁存，阈值类仍属组态非法并锁存 *)
_bMeasBad := (fEnergy <> fEnergy) OR (fDisp <> fDisp) OR (fPressure <> fPressure);          // 实测 NaN 自反判（单列出口） / Measured NaN tests, separate outlet
_bThBad   := (fEnergyLo <> fEnergyLo) OR (fEnergyHi <> fEnergyHi)                          // 能量窗 NaN 判 / Energy envelope NaN tests
          OR (fDispLo <> fDispLo) OR (fDispHi <> fDispHi)                                  // 位移窗 NaN 判 / Displacement envelope NaN tests
          OR (fPressLo <> fPressLo) OR (fPressHi <> fPressHi);                             // 压力窗 NaN 判 / Pressure envelope NaN tests
_bNonFin  := _bMeasBad OR _bThBad;                                                         // 非有限汇总（诊断口径保留） / Aggregated non-finite flag
_bCfgBad  := (fEnergyLo >= fEnergyHi) OR (fDispLo >= fDispHi) OR (fPressLo >= fPressHi)    // 六阈值双侧几何闸（倒置即恒 NG） / Six-threshold geometry gate
          OR _bThBad;                                                                      // 仅阈值类非有限并入组态非法 / Threshold non-finite folded into config
rtEval(CLK := bEval);                                                              // 评估沿，每拍必调（R228A） / Evaluation edge, every scan
rtReset(CLK := bReset);                                                            // 复位沿，每拍必调 / Reset edge, every scan

(* —— 段 1：单拍量预清零（锁存量 _bNg1/_bNg2/_bNg3/_bAnyNg/_eCause 不入清单，R107） —— *)
bEvalDone := FALSE;         // 评估完成脉冲每拍预清 / Eval-done pulse preset
bError    := FALSE;         // 故障标志每拍预清（R45 配对） / Error flag preset
_bE1      := FALSE;         // 本次能量 NG 预清 / Energy NG preset
_bE2      := FALSE;         // 本次位移 NG 预清 / Displacement NG preset
_bE3      := FALSE;         // 本次压力 NG 预清 / Pressure NG preset
_nNgCnt   := 0;             // 越窗计数预清 / NG count preset

(* —— 段 2：复位沿（唯一清锁存路径） —— *)
IF rtReset.Q THEN
    _bNg1   := FALSE;                       // 清能量 NG 锁存 / Clear energy NG latch
    _bNg2   := FALSE;                       // 清位移 NG 锁存 / Clear displacement NG latch
    _bNg3   := FALSE;                       // 清压力 NG 锁存 / Clear pressure NG latch
    _bAnyNg := FALSE;                       // 清任一路 NG 锁存 / Clear any-NG latch
    _eCause := E_DL_TwmCause.eNone;         // 清成因 / Clear cause
    IF _eState = E_DL_TwmState.eFault THEN
        _eState := E_DL_TwmState.eIdle;     // 故障相迁出（R228B） / Leave fault phase
    END_IF
END_IF

(* —— 段 3：组态闸（闸门故障不得记成焊点 NG，故不置任何通道位） —— *)
IF _bCfgBad THEN
    _eState := E_DL_TwmState.eFault;        // 入故障相 / Enter fault phase
    _eCause := E_DL_TwmCause.eCfgIllegal;   // 归因：组态非法 / Cause: illegal configuration
END_IF

(* —— 段 3b：实测 NaN 单列出口（当拍跳过评估，不锁存、不动任何通道位，v1.0.1） —— *)
IF rtEval.Q AND _bMeasBad THEN
    _eCause := E_DL_TwmCause.eMeasBad;      // 归因：实测值 NaN / Cause: measured NaN
END_IF

(* —— 段 4：评估沿——三路独立双侧包络判定（单点写入锁存，避免同拍抹除，R187） —— *)
IF rtEval.Q AND (NOT _bCfgBad) AND (NOT _bMeasBad) THEN
    _bE1 := (fEnergy < fEnergyLo) OR (fEnergy > fEnergyHi);        // 能量双侧越窗（下限也要查） / Energy outside both bounds
    _bE2 := (fDisp < fDispLo) OR (fDisp > fDispHi);                // 位移双侧越窗 / Displacement outside both bounds
    _bE3 := (fPressure < fPressLo) OR (fPressure > fPressHi);      // 压力双侧越窗 / Pressure outside both bounds
    IF _bE1 THEN
        _bNg1 := TRUE;                                             // 能量 NG 锁存 / Latch energy NG
    END_IF
    IF _bE2 THEN
        _bNg2 := TRUE;                                             // 位移 NG 锁存 / Latch displacement NG
    END_IF
    IF _bE3 THEN
        _bNg3 := TRUE;                                             // 压力 NG 锁存 / Latch pressure NG
    END_IF
    IF _bE1 THEN
        _nNgCnt := _nNgCnt + 1;                                    // 计数 +1（USINT 上限 5 远够） / Count up, USINT is ample
    END_IF
    IF _bE2 THEN
        _nNgCnt := _nNgCnt + 1;
    END_IF
    IF _bE3 THEN
        _nNgCnt := _nNgCnt + 1;
    END_IF
    IF _nNgCnt > 0 THEN
        _bAnyNg := TRUE;                                           // 累计任一 NG 锁存 / Latch the accumulated any-NG
        IF _nNgCnt = 1 THEN
            IF _bE1 THEN
                _eCause := E_DL_TwmCause.eEnergyNg;                // 归因：唯一越窗=能量 / Cause: energy is the only channel
            ELSIF _bE2 THEN
                _eCause := E_DL_TwmCause.eDispNg;                  // 归因：唯一越窗=位移 / Cause: displacement is the only channel
            ELSE
                _eCause := E_DL_TwmCause.ePressNg;                 // 归因：唯一越窗=压力 / Cause: pressure is the only channel
            END_IF
        ELSE
            _eCause := E_DL_TwmCause.eMultiNg;                     // 归因：多路同时越窗（不强行挑一条） / Cause: multiple channels, no forced pick
        END_IF
    END_IF
    bEvalDone := TRUE;                                             // 单拍评估完成 / Single-scan evaluation done
    IF _eState = E_DL_TwmState.eIdle THEN
        _eState := E_DL_TwmState.eRun;                             // 首次评估后进入运行相 / First evaluation enters run phase
    END_IF
END_IF

(* —— 段 5：相位机（ENUM 全成员显式标签 + ELSE 兜底，R128） —— *)
CASE _eState OF

E_DL_TwmState.eIdle:
    IF _bCfgBad THEN                                            // 出口 1：组态非法 / Illegal configuration
        _eState := E_DL_TwmState.eFault;
    ELSIF rtEval.Q THEN                                         // 出口 2：首次评估沿 / First evaluation edge
        _eState := E_DL_TwmState.eRun;
    END_IF

E_DL_TwmState.eRun:
    IF _bCfgBad THEN                                            // 出口 1：组态转非法 / Configuration went illegal
        _eState := E_DL_TwmState.eFault;
    ELSIF rtReset.Q THEN                                        // 出口 2：复位回等待相 / Reset back to idle
        _eState := E_DL_TwmState.eIdle;
    END_IF

E_DL_TwmState.eFault:
    IF rtReset.Q AND (NOT _bCfgBad) THEN                        // 出口：复位且组态已合法才迁出（R228B） / Reset with legal config
        _eState := E_DL_TwmState.eIdle;
    END_IF

ELSE
    _eCause := E_DL_TwmCause.ePhaseBad;                         // 归因：非法相位 / Cause: illegal phase
    _eState := E_DL_TwmState.eFault;                            // 强拉故障相 / Force fault phase
    bError  := TRUE;                                            // 故障标志 / Error flag

END_CASE

(* —— 段 6：出口单点映射（三路独立 + 掩码同源；名实双出口 R191） —— *)
bEnergyNg := _bNg1;                                             // 能量 NG 出口 / Energy NG outlet
bDispNg   := _bNg2;                                             // 位移 NG 出口 / Displacement NG outlet
bPressNg  := _bNg3;                                             // 压力 NG 出口 / Pressure NG outlet
bAnyNg    := _bAnyNg;                                           // 任一路 NG 出口（锁存累计） / Any-NG outlet
nNgMask   := 16#00;                                             // 掩码每拍重建（由三路 BOOL 派生，不独立维护） / Mask rebuilt from the three flags
IF _bNg1 THEN
    nNgMask := nNgMask OR DL_TWM_MASK_E;                        // bit0 能量 / bit0 energy
END_IF
IF _bNg2 THEN
    nNgMask := nNgMask OR DL_TWM_MASK_D;                        // bit1 位移 / bit1 displacement
END_IF
IF _bNg3 THEN
    nNgMask := nNgMask OR DL_TWM_MASK_P;                        // bit2 压力 / bit2 pressure
END_IF
bError  := _bAnyNg OR (_eState = E_DL_TwmState.eFault);         // 故障标志 = 任一路 NG 或组态故障 / Error = any NG or config fault
eState  := _eState;                                             // 状态出口 / State outlet
eCause  := _eCause;                                             // 成因出口 / Cause outlet

END_FUNCTION_BLOCK
